(* IEC 61131-3 sources: daoli-st-library/DL_Base (part 9) *)

(* ---- FB_DL_AlarmShelveMgmt.st ---- *)
(*==============================================================================
 * 组件名称 (Component)  : FB_DL_AlarmShelveMgmt
 * 所属子库 (Sublibrary) : DL_Base
 * 当前版本 (Version)    : 1.0.0
 * 兼容性   (Platform)   : CODESYS 3.5 / TwinCAT 3 / 汇川 InoProShop / Machine Expert
 *                         仅依赖 Standard.library（TON / R_TRIG），零厂商方言
 * 来源标签 (Source)     : isa-18.2（T2-8 报警管理族本体：搁置 Shelving 生命周期）
 * 功能描述 (Function)   : ISA-18.2 报警搁置管理状态机：申请沿 -> 搁置生效（带时限）->.
 *                         时限到期自动解除；人工解除沿即时恢复。搁置申请 / 人工解除 /
 *                         自动解除三类事件写入 4 条深度环形审计台账（带全局序号）。
 * 分工互引 (Boundary)   : FB_DL_AlarmFloodLimiter 做报警**限流**（抑制短时洪泛），
 *                         本件做**搁置**（操作员主动、有时限、必须留痕）；两者语义
 *                         不同不可互代（限流不改报警状态，搁置改报警可见性）。
 *                         报警本体与优先级归 FB_DL_AlarmManager。
 * 边界与语义披露 (Boundary disclosure) :
 *   1) 搁置时限 tShelveDur <= T#0S 属组态非法：拒绝进入搁置并置故障级，锁存至
 *      复位沿 + 组态改对（R152 解除路径自证可达）。
 *   2) 同拍「申请 + 解除」：解除优先（安全侧），申请作废不入台账。
 *   3) 只允许单报警搁置（uAlarmId 单槽）：多报警并发搁置由上层按报警号各实例化
 *      一份本件（组合优于在件内做动态表，避免变长容器）。
 *   4) 审计台账 4 条环形：写满覆盖最旧并置一次性信息码；写指针显式归零，不做越界写。
 *   5) 搁置状态在 bEnable 拉低时**保持**（不静默解除）：失能不是解除条件，
 *      解除只能来自人工解除沿或时限到期（避免上位机失能导致报警被永久藏起来）。
 * 故障码表 (Error codes) :
 *   16#0001_03FE [故障级] 搁置时限组态非法（<= T#0S），拒绝进入搁置
 *                 反证：拒绝搁置与「操作员没申请」输出组合完全相同，无码不可区分。
 *   16#0001_04FA [信息级] 搁置生效（申请沿受理并入台账）
 *                 反证：bShelved 只表达状态，无法承载「何时由谁申请」的事件事实。
 *   16#0001_04FB [信息级] 时限到期自动解除（旁路被时限收割）
 *                 反证：自动解除与人工解除对外同形（都退出搁置），仅事件种类不同。
 *   16#0001_04FC [信息级] 审计台账环形已回卷（最旧条目被覆盖）
 *                 反证：回卷后 nAuditCount 恒为 4，与「恰好写满」输出组合相同。
 * 码位总账 (Code ledger) : 16#0001_03FE 用 ｜ 16#0001_04FA / 04FB / 04FC 用
 * 依赖     (Depends)    : 无 DL_ 内部依赖；Standard.library: TON / R_TRIG
 * 红线自检 (Redline)    : R1 ✓ 零全局变量 ｜ R2 ✓ 零 %I/%Q ｜ R3 ✓ 纯 IEC 61131-3
 *                         R4 ✓ 时限判零 / 环形显式回卷无越界 ｜ R5 ✓ 全变量双语同行注释
 *                         R6 ✓ 三态 ENUM + CASE + ELSE 兜底 ｜ R7 ✓ 三沿一计时最前部无条件刷新
 * 修订历史 (Revision)   : 2026-11-22  v1.0.0  首版入库（R69 构建轮 · 批 2 · N6）
 *============================================================================*)

(*-----------------------------------------------------------------------------
 * 枚举: E_DL_ShelveState / E_DL_ShelveEvt（归属 DL_Base，与 FB_DL_AlarmShelveMgmt 同文件）
 *----------------------------------------------------------------------------*)
TYPE E_DL_ShelveState :
(
    eIdle    := 0,    // 未搁置：报警正常可见 / Not shelved, the alarm stays visible
    eShelved := 10,   // 搁置生效：时限窗计时 / Shelved, the time window runs
    eFault   := 99    // 组态故障：拒绝一切新搁置 / Config fault, new shelving refused
);
END_TYPE

TYPE E_DL_ShelveEvt :
(
    eNone     := 0,   // 无事件（空槽哨兵）/ No event, empty slot sentinel
    eApply    := 1,   // 申请搁置 / Shelving applied
    eRelCmd   := 2,   // 人工解除 / Released by the operator
    eRelTime  := 3    // 时限自动解除 / Released by the time window
);
END_TYPE

(*==============================================================================
 * 功能块: FB_DL_AlarmShelveMgmt
 * 调用约定: 每个扫描周期无条件调用一次；bShelveReq / bUnshelveReq 为上升沿语义。
 *============================================================================*)
FUNCTION_BLOCK FB_DL_AlarmShelveMgmt
VAR_INPUT
    bShelveReq    : BOOL;                  // 搁置申请，上升沿生效 / shelving request, rising edge
    bUnshelveReq  : BOOL;                  // 人工解除，上升沿生效 / manual release, rising edge
    uAlarmId      : UINT := 0;             // 被搁置报警号 [号]，随事件入台账 / alarm id logged with each event
    tShelveDur    : TIME := T#30M;         // 搁置时限 [s]，<= T#0S 组态非法 / shelving duration [s]
    bEnable       : BOOL := TRUE;          // 使能；FALSE 只冻结新申请，不解除已搁置 / enable, FALSE freezes new requests only
    bReset        : BOOL;                  // 上升沿：清组态故障锁存 / rising edge clears the config latch
END_VAR
VAR_OUTPUT
    bShelved      : BOOL;                  // 搁置生效中（报警可被 HMI 隐藏）/ shelving active
    tElapsed      : TIME;                  // 已搁置时长 [s] / elapsed shelving time [s]
    tRemain       : TIME;                  // 剩余搁置时长 [s] / remaining shelving time [s]
    bExpired      : BOOL;                  // 本拍时限到期（单拍脉冲）/ window expired, single scan
    nAuditCount   : INT;                   // 台账有效条数 [条]，0..4 / valid ledger entries
    bAuditWrapped : BOOL;                  // 台账已回卷覆盖 / ledger wrapped
    eLastEvt      : E_DL_ShelveEvt;        // 最近事件种类 / kind of the most recent event
    uLastEvtSeq   : UDINT;                 // 最近事件全局序号 [号] / global sequence of the last event
    auLedgerAlarm : ARRAY[0..3] OF UINT;   // 台账报警号环形副本 [号] / ledger alarm id ring copy
    aLedgerEvt    : ARRAY[0..3] OF E_DL_ShelveEvt; // 台账事件种类环形副本 / ledger event kind ring copy
    bError        : BOOL;                  // 故障标志（组态锁存）/ fault flag
    uErrorId      : UDINT;                 // 故障码，0 = 无故障 / error code, 0 = none
    eState        : E_DL_ShelveState;      // 当前状态（供 HMI 诊断）/ current state
END_VAR
VAR
    fbTrigReq     : R_TRIG;                // 申请沿检测实例 / request edge detector
    fbTrigRel     : R_TRIG;                // 解除沿检测实例 / release edge detector
    fbTrigReset   : R_TRIG;                // 复位沿检测实例 / reset edge detector
    tonShelve     : TON;                   // 搁置时限计时实例 / shelving window timer
    eStateInt     : E_DL_ShelveState;      // 主状态机内部当前态 / internal state
    bDurBad       : BOOL;                  // 本拍时限组态非法 / duration illegal this scan
    bCfgLatch     : BOOL;                  // 组态锁存（复位沿 + 组态改对解除）/ config latch
    bShelveOn     : BOOL;                  // 搁置驻留标志（驱动 TON.IN）/ shelving dwell flag driving TON.IN
    bExpiredT     : BOOL;                  // 到期脉冲内部副本（单拍）/ internal expired pulse
    aeEvtInt      : ARRAY[0..3] OF E_DL_ShelveEvt; // 台账事件种类（内部）/ ledger event kind ring, internal
    auiAlarmInt   : ARRAY[0..3] OF UINT;   // 台账报警号（内部）/ ledger alarm id ring, internal
    nWriteIdx     : INT;                   // 台账写指针 [0..3] / ledger write pointer
    uEvtTotal     : UDINT;                 // 累计事件总数 [件]（回卷判据）/ total events ever
    uSeqInt       : UDINT;                 // 全局序号计数器 [号]，饱和 / saturating sequence counter
    bWrapCoded    : BOOL;                  // 回卷事件码已发（一次性）/ wrap event already coded
    uTargetInt    : UINT;                  // 入场报警号内部副本 [号] / internal alarm id copy
    eLastEvtInt   : E_DL_ShelveEvt;        // 最近事件种类内部副本 / internal last event kind
    uLastSeqInt   : UDINT;                 // 最近事件序号内部副本 / internal last sequence
    bErrorInt     : BOOL;                  // 本拍故障置位累加 / fault set accumulator
    bFirstScan    : BOOL := TRUE;          // 上电首扫标志 / first-scan flag
END_VAR
VAR CONSTANT
    DL_AS_DEPTH   : INT := 4;              // 台账环形深度 [条] / ledger ring depth
    DL_AS_SEQ_MAX : UDINT := 16#FFFF_FFFE; // 序号饱和上界 [号] / sequence saturation bound
END_VAR

METHOD WriteAudit
VAR_INPUT
    eEvt : E_DL_ShelveEvt;          // 待写事件种类 / event kind to be written
END_VAR
VAR
    nSlot : INT;                    // 本次写入槽位 [0..3] / slot index of this write
END_VAR

nSlot := nWriteIdx;                              // 取当前写指针 / take the current pointer
aeEvtInt[nSlot]    := eEvt;                      // 事件种类入账 / event kind into the ledger
auiAlarmInt[nSlot] := uTargetInt;                // 报警号入账 / alarm id into the ledger
IF uSeqInt < DL_AS_SEQ_MAX THEN
    uSeqInt := uSeqInt + 1;                      // 序号推进（饱和）/ advance the sequence, saturating
END_IF
uLastSeqInt   := uSeqInt;                        // 最近序号留影 / snapshot the sequence
eLastEvtInt   := eEvt;                           // 最近事件种类留影 / snapshot the kind
uEvtTotal     := uEvtTotal + 1;                  // 累计事件推进（回卷判据）/ total events up
nWriteIdx     := nWriteIdx + 1;                  // 写指针推进 / advance the pointer
IF nWriteIdx >= DL_AS_DEPTH THEN
    nWriteIdx := 0;                              // 显式回卷（IF 等价，禁 MOD 方言）/ explicit wrap
END_IF

END_METHOD

(*------------------------------------------------------------------------------
 * 段 1｜无条件刷新区（红线 R7）：三沿一计时位于主体最前部
 *      Unconditional refresh: three edges and one timer at the very top
 *-----------------------------------------------------------------------------*)
fbTrigReq(CLK := bShelveReq);
fbTrigRel(CLK := bUnshelveReq);
fbTrigReset(CLK := bReset);
tonShelve(IN := bShelveOn, PT := tShelveDur);   // IN 用内部驻留标志，禁挂外部引脚原值 / driven by the internal dwell flag

(* 段 2｜上电首扫：台账槽位显式落哨兵 / first-scan init *)
IF bFirstScan THEN
    FOR nWriteIdx := 0 TO (DL_AS_DEPTH - 1) DO
        aeEvtInt[nWriteIdx] := E_DL_ShelveEvt.eNone;   // 空槽哨兵 / empty slot sentinel
    END_FOR
    nWriteIdx   := 0;
    uEvtTotal   := 0;
    uSeqInt     := 0;
    eStateInt   := E_DL_ShelveState.eIdle;
    bFirstScan  := FALSE;
END_IF

(* 段 3｜每拍预清（FB32-1）：单拍标志，禁入锁存 / per-scan preset *)
bErrorInt := FALSE;
bExpiredT := FALSE;

(*------------------------------------------------------------------------------
 * 段 4｜组态域闸：时限 <= 0 非法，锁存至复位沿 + 组态改对（R152 自证可达）
 *      Config gate on the shelving duration with the reachable clear path
 *-----------------------------------------------------------------------------*)
bDurBad := (tShelveDur <= T#0S);
IF bDurBad THEN
    bCfgLatch := TRUE;
END_IF
IF fbTrigReset.Q AND (NOT bDurBad) THEN
    bCfgLatch := FALSE;              // 组态锁存解除 / config latch cleared
    uErrorId  := 16#0000_0000;       // 码位随解除归零 / code cleared with the latch
END_IF
IF bCfgLatch THEN
    uErrorId  := 16#0001_03FE;       // 故障级：时限组态非法 / fault: illegal duration
    bErrorInt := TRUE;               // R45 配对 / paired with the code
    eStateInt := E_DL_ShelveState.eFault;
    bShelveOn := FALSE;              // 迁相补清：故障打断搁置即断计时 / timing dropped on migration
END_IF

(*------------------------------------------------------------------------------
 * 段 5｜主状态机（红线 R6）：ENUM + CASE + ELSE 兜底
 *      同拍竞态（R275）：eShelved 相内先消化解除沿，再消化时限到期
 *-----------------------------------------------------------------------------*)
CASE eStateInt OF

    E_DL_ShelveState.eIdle:
        (* 同拍「申请 + 解除」：解除优先（安全侧），申请作废不入台账 *)
        IF bEnable AND (NOT bCfgLatch) AND fbTrigReq.Q AND (NOT fbTrigRel.Q) THEN
            uTargetInt := uAlarmId;                       // 报警号留影 [号] / snapshot the alarm id
            bShelveOn  := TRUE;                           // 起计时 / start the window
            uErrorId   := 16#0000_0000;                   // 新一轮开始，旧事件码回落 / previous event codes fall back
            WriteAudit(eEvt := E_DL_ShelveEvt.eApply);    // 入台账 / write the audit entry
            eStateInt  := E_DL_ShelveState.eShelved;
        END_IF

    E_DL_ShelveState.eShelved:
        IF fbTrigRel.Q THEN
            bShelveOn  := FALSE;                          // 人工解除即时生效 / manual release is immediate
            uTargetInt := uAlarmId;
            WriteAudit(eEvt := E_DL_ShelveEvt.eRelCmd);
            eStateInt  := E_DL_ShelveState.eIdle;
        ELSIF tonShelve.Q THEN
            bShelveOn  := FALSE;                          // 时限到期自动解除 / auto release on expiry
            uTargetInt := uAlarmId;
            uErrorId   := 16#0001_04FB;                   // 信息级：时限自动解除 / info: auto released
            bExpiredT  := TRUE;                           // 单拍到期脉冲 / single-scan expired pulse
            WriteAudit(eEvt := E_DL_ShelveEvt.eRelTime);
            eStateInt  := E_DL_ShelveState.eIdle;
        END_IF

    E_DL_ShelveState.eFault:
        IF fbTrigReset.Q AND (NOT bDurBad) THEN
            bCfgLatch := FALSE;                           // 解除路径自证可达 / clear path reachable
            uErrorId  := 16#0000_0000;
            eStateInt := E_DL_ShelveState.eIdle;
        END_IF

    ELSE
        (* 非法状态拦截 / illegal state interception *)
        eStateInt := E_DL_ShelveState.eFault;
        uErrorId  := 16#0001_03FE;
        bErrorInt := TRUE;

END_CASE;

(*------------------------------------------------------------------------------
 * 段 6｜输出单一出口（范式 P-05）：搁置位只由状态派生一次
 *      Single output exit: the shelved bit derives from the state exactly once
 *-----------------------------------------------------------------------------*)
bShelved     := (eStateInt = E_DL_ShelveState.eShelved);
tElapsed     := tonShelve.ET;                            // 已搁置时长 [s] / elapsed time
IF tShelveDur > tonShelve.ET THEN
    tRemain  := tShelveDur - tonShelve.ET;               // 剩余时长 [s] / remaining time
ELSE
    tRemain  := T#0S;                                    // 已到期：剩余 0 [s] / expired, zero remaining
END_IF
bExpired     := bExpiredT;                               // 单拍脉冲统一出口 / unified single-scan exit
bAuditWrapped := (uEvtTotal > UDINT#4);                  // 回卷事实量（常驻，与事件码分离）/ wrapped standing fact
IF bAuditWrapped AND (NOT bWrapCoded) THEN
    uErrorId   := 16#0001_04FC;                          // 信息级：台账回卷（一次性）/ info: wrapped once
    bWrapCoded := TRUE;
END_IF
IF fbTrigReset.Q AND (NOT bCfgLatch) THEN
    uErrorId   := 16#0000_0000;                          // 信息码随复位沿回落 / info codes fall back
    bWrapCoded := FALSE;
END_IF
IF UDINT_TO_DINT(uEvtTotal) < DINT#4 THEN
    nAuditCount := DINT_TO_INT(UDINT_TO_DINT(uEvtTotal));
ELSE
    nAuditCount := DL_AS_DEPTH;                          // 深度即上限 [条] / depth is the cap
END_IF
eLastEvt    := eLastEvtInt;
uLastEvtSeq := uLastSeqInt;
FOR nWriteIdx := 0 TO (DL_AS_DEPTH - 1) DO
    aLedgerEvt[nWriteIdx]   := aeEvtInt[nWriteIdx];      // 台账副本直出 / ledger copy out
    auLedgerAlarm[nWriteIdx] := auiAlarmInt[nWriteIdx];
END_FOR
bError := bErrorInt OR bCfgLatch;
eState := eStateInt;

(*------------------------------------------------------------------------------
 * 私有方法: WriteAudit —— 审计台账唯一写入点（指针 / 序号 / 计数三记账）
 *      Private method: the single audit write entry
 *      调用约定: 仅在本件主体 CASE 内调用，无阻塞、无 METHOD 内跨周期驻留
 *-----------------------------------------------------------------------------*)

END_FUNCTION_BLOCK

(* ---- FB_DL_BitArrayChangeWatch.st ---- *)
(*==============================================================================
 * 组件名称 (Component)  : FB_DL_BitArrayChangeWatch
 * 所属子库 (Sublibrary) : DL_Base
 * 归属目录 (Directory)  : C:\Library\DL_Base
 * 当前版本 (Version)    : 1.0.1
 * 组件分类 (Category)   : 功能块（FUNCTION_BLOCK）· 位图变化监视 · 状态机
 * 兼容性   (Platform)   : CODESYS 3.5 / TwinCAT 3 / 汇川 InoProShop / 施耐德
 *                         Machine Expert；仅用 Standard.library 的 R_TRIG 与位运算
 * 功能一句话 (Summary)  : 逐拍监视 DWORD 数组位图的位级变化，输出本拍变化掩码、
 *                         变化位数、首个变化位绝对位号，并累计跳变次数与判稳标志。
 * 功能描述 (Function)   : 上位机只显示「有变化」时不定位，接触不良的端子表现为
 *                         某一位反复抖动，必须单独统计跳变位数才能定位到端子与
 *                         线号。本件把「本拍变化」与「累计抖动」分开输出：变化掩码
 *                         给 HMI 做位闪烁，跳变累计给维修工排出最脏的位。
 * 与既有件边界 (Boundary): FC_DL_DualEdgeTrig 做单信号的边沿检测；FB_DL_SignalDebounce
 *                         做单信号滤波；本件做整组位图的位级变化统计，三者正交。
 * 设计要点 (Key notes)  : ① 复位沿检测实例在状态机之外无条件刷新，绝不放进分支；
 *                         ② 首拍只装载不复位跳变计数，避免上电瞬间误报全部位跳动；
 *                         ③ 跳变累计饱和不回绕：回绕会把抖动最严重的位算成最干净的位；
 *                         ④ 掉使能只清变化族，不清跳变累计，诊断证据不因停机而丢失；
 *                         ⑤ 快照赋值放在输出之后，保证下一拍才参与比较；
 *                         ⑥ 位扫描与首变位查找合并为一趟循环，避免两趟扫描的节拍差。
 * 开源溯源 (Origin)     : 来源标签 lgf-bitlogic。LGF 为免费闭源发布的公开函数库手册，
 *                         本件仅借鉴其位逻辑组把「单点位测试」与「批量监视」并列的
 *                         分类位置；许可证按其发布方条款仅作分类参考，变化检测算法、
 *                         跳变统计与饱和策略全部自有，属 clean-room 独立实现。
 * 码位说明 (Codes)      : 信息级 16#0001_012D 字数上限钳位 ｜ 16#0001_012E 判稳拍数
 *                         钳位 ｜ 16#0001_012F 跳变累计饱和；
 *                         故障级 16#0001_021A 字数小于一（组态错，锁存）｜
 *                         16#0001_021B 非法状态兜底。故障级码只在本件使用，
 *                         与全库已占码求差为空。
 * 依赖说明 (Depends)    : 无 DL_ 内部依赖；仅 Standard.library 的 R_TRIG 与
 *                         SHL / XOR / INT_TO_UDINT / UDINT_TO_INT。
 * 调用约定 (Call rules): 每扫描周期无条件调用一次；bEnable 为假时输出变化族清零，
 *                         跳变累计保持，恢复使能后继续累加。
 * 红线自检 (Redline)    : 零全局变量表依赖 ｜ 零外部变量声明 ｜ 零物理地址
 *                         纯 IEC 61131-3 ｜ 数组下标先钳位后使用 ｜ 无除法
 *                         状态机三成员全覆盖并带兜底 ｜ 边沿实例在分支外刷新
 * 修订历史 (Revision)   : 2026-11-15  v1.0.0  首版入库（Round 12 · 位图变化监视）
 *                         2026-11-15  v1.0.1  终审定点修复 A-D03：掉使能回空闲的判据补
 *                         「当前不在故障态」前置条件，杜绝使能为假时抢走复位上升沿
 *                         导致故障不可复位（eFault 主体整拍被跳过，边沿一拍即失）
 *============================================================================*)

(*-----------------------------------------------------------------------------
 * 枚举: E_DL_BitWatchState（归属 DL_Base，与 FB_DL_BitArrayChangeWatch 同文件）
 * 含义: 位图监视主状态。编号 0 起跳、段间隔 10，便于后续插态。
 *----------------------------------------------------------------------------*)
TYPE E_DL_BitWatchState :
(
    eIdle     := 0,      // 空闲：装载快照并清零变化族，等待使能 / Idle, snapshot loaded when enabled
    eSampling := 10,     // 采样：逐字比对、位统计、跳变累计与判稳 / Sampling, compare and accumulate every cycle
    eFault    := 99      // 故障：组态错锁存，输出冻结，复位沿退出 / Latched configuration fault, outputs frozen
);
END_TYPE

(*==============================================================================
 * 拍序示意 (Cycle sequence)：
 *   第 1 拍  空闲态装载上拍快照，本拍不比较，故不产生跳变
 *   第 2 拍  采样态比较本拍与上拍，异或结果即变化掩码，同时累计跳变位数
 *   第 3 拍  若连续无变化拍数达到判稳门限，判稳标志置真
 *   第 4 拍  快照更新为第 3 拍的位图，第 5 拍起以新快照为基准
 *   跳变累计只在采样态累加，首拍装载与掉使能期间一律不动
 *============================================================================*)

FUNCTION_BLOCK FB_DL_BitArrayChangeWatch
VAR_INPUT
    bEnable       : BOOL;                          // 使能，为假时变化族清零并退出采样 / Enable, clears the change family when false
    bReset        : BOOL;                          // 上升沿复位跳变累计与判稳计时 / Rising edge resets toggle count and settle timer
    nWordCount    : INT := 1;                      // 监视字数 [个]，域 1 到 8，越界钳位 / Watched word count, 1 to 8, clamped
    auWatch       : ARRAY[1..8] OF DWORD;          // 当前位图快照，位 0 在最低位 [位串] / Current bitmap snapshot, bit zero is the lowest bit
    nSettleCycles : INT := 2;                      // 判稳所需连续无变化拍数 [拍]，域 1 到 100 / Cycles required to declare steady, 1 to 100
END_VAR
VAR_OUTPUT
    auChangeMask  : ARRAY[1..8] OF DWORD;          // 本拍变化位掩码，按字对齐，未监视的字为零 [位串] / Per word change mask of this cycle
    nChangeBits   : INT;                           // 本拍变化位总数，逐字位计数之和 [位] / Total changed bits this cycle
    nFirstBit     : INT;                           // 首个变化位绝对位号，负一表示本拍无变化 [bit] / First changed absolute bit, minus one when none
    uToggleCount  : UDINT;                         // 累计跳变位数，由复位上升沿清零 [位次] / Accumulated toggled bits, cleared by the reset edge
    bSteady       : BOOL;                          // 连续无变化拍数达到门限为真 / No change for the settle window
    eState        : E_DL_BitWatchState;            // 主状态机当前状态，供 HMI 诊断 / Current state of the main state machine
    bError        : BOOL;                          // 故障级锁存，仅字数小于一与非法状态置位 / Latched fault, only set by the two fault codes
    uErrorId      : UDINT;                         // 事件码，0 表示无事件 / Event code, zero means none
END_VAR
VAR
    auPrev        : ARRAY[1..8] OF DWORD;          // 上拍快照，跨周期保持 [位串] / Previous snapshot kept across cycles
    auXor         : ARRAY[1..8] OF DWORD;          // 本拍异或结果 [位串] / XOR result of this cycle
    fbTrigReset   : R_TRIG;                        // 复位沿检测实例，在状态机之外无条件刷新 / Reset edge detector refreshed outside the state machine
    eStateInt     : E_DL_BitWatchState := E_DL_BitWatchState.eIdle; // 内部状态，对外经 eState 输出 / Internal state exported through eState
    bFirstScan    : BOOL := FALSE;                 // 首拍装载完成标志，初值假表示尚未装载 / First scan loaded flag, false means not yet loaded
    nWordClamped  : INT;                           // 钳位后字数 [个] / Clamped word count
    nSettleUse    : INT;                           // 生效判稳拍数 [拍] / Effective settle cycles
    nSteadyCnt    : INT;                           // 已连续无变化拍数 [拍] / Cycles already steady
    uWeight       : UDINT;                         // 单拍位计数中间量 [位] / Population count intermediate
    nBitScan      : INT;                           // 位扫描索引，0 到 31 [bit] / Bit scan index, 0 to 31
    nIdx          : INT;                           // 字下标遍历索引 [索引] / Word loop index
    nGuard        : DINT;                          // 循环守卫计数，防字循环失控 [次] / Loop guard counter for the word loop
    bAnyChange    : BOOL;                          // 本拍是否发生变化 / Any change this cycle
    bParamClamped : BOOL;                          // 参数被钳位标记，故障态退出判据之一 / Parameter clamped flag, also gates the fault exit
END_VAR
VAR CONSTANT
    DL_WORD_MAX   : INT := 8;                          // 字数上限 [个] / Word count limit
    DL_BIT_WORD   : INT := 32;                         // 单字位宽 [bit] / Bits per word
    DL_GUARD_MAX  : DINT := 64;                        // 循环守卫上限，远大于字数上限故正常不触发 [次] / Loop guard limit, never reached in normal operation
    DL_I_W        : INT := 1;                          // 数组首下标 [索引] / First array index
    DL_SETTLE_MIN : INT := 1;                          // 判稳拍数下限 [拍] / Lower settle bound
    DL_SETTLE_MAX : INT := 100;                        // 判稳拍数上限，同时兼作稳定计数饱和值 [拍] / Upper settle bound, also saturates the steady counter
    DL_TOGGLE_MAX : UDINT := 16#FFFF_FFFE;             // 跳变累计饱和值，禁止回绕 [位次] / Saturation value of the toggle counter, no wrap around
END_VAR

(*------------------------------------------------------------------------------
 * 段 1｜复位沿检测（红线）：实例在状态机之外每拍无条件刷新
 *      Reset edge detector, refreshed unconditionally outside the state machine
 *-----------------------------------------------------------------------------*)
fbTrigReset(CLK := bReset);

(*------------------------------------------------------------------------------
 * 段 2｜事件码刷新与参数钳位（边界 B1/B2）
 *      Event code refresh and parameter clamping
 *      未锁存故障时每拍先清码，保证事件码是「本拍事件」而不是陈年旧码
 *-----------------------------------------------------------------------------*)
IF NOT bError THEN
    uErrorId := 16#0000_0000;
END_IF

nWordClamped := nWordCount;
IF nWordClamped < DL_I_W THEN
    nWordClamped  := DL_I_W;
    bParamClamped := TRUE;
    bError        := TRUE;
    uErrorId      := 16#0001_021A;   // 组态错：字数小于一，属数组域非法
ELSE
    bParamClamped := FALSE;
    IF nWordClamped > DL_WORD_MAX THEN
        nWordClamped  := DL_WORD_MAX;
        bParamClamped := TRUE;
        IF uErrorId = 16#0000_0000 THEN
            uErrorId := 16#0001_012D;   // 字数超限，已钳位到上限并照常服务
        END_IF
    END_IF
END_IF

nSettleUse := nSettleCycles;
IF nSettleUse < DL_SETTLE_MIN THEN
    nSettleUse := DL_SETTLE_MIN;
    IF uErrorId = 16#0000_0000 THEN
        uErrorId := 16#0001_012E;   // 判稳拍数过小，已钳到下限
    END_IF
ELSIF nSettleUse > DL_SETTLE_MAX THEN
    nSettleUse := DL_SETTLE_MAX;
    IF uErrorId = 16#0000_0000 THEN
        uErrorId := 16#0001_012E;   // 判稳拍数过大，已钳到上限
    END_IF
END_IF

(*------------------------------------------------------------------------------
 * 段 3｜复位沿副作用：清跳变累计与判稳计时，故障退出由状态机自行处理
 *      Reset side effects: clear the toggle count and the settle timer
 *-----------------------------------------------------------------------------*)
IF fbTrigReset.Q AND (eStateInt <> E_DL_BitWatchState.eFault) THEN
    uToggleCount := 0;
    nSteadyCnt   := 0;
    bSteady      := FALSE;
END_IF

(*------------------------------------------------------------------------------
 * 段 4｜掉使能统一回空闲（边界 B3）：跳变累计不清，诊断证据保留
 *      Disable forces idle, the toggle counter is deliberately preserved
 *      故障态不放行：eFault 的复位沿判据必须每拍都有机会执行，若在此处无条件
 *      改写为 eIdle，CASE 只会进 eIdle 分支，故障态主体整拍被跳过、复位上升沿
 *      一拍即失（现场「停机后按复位无效」的典型成因）
 *      The fault phase is excluded so that its reset edge is never skipped
 *-----------------------------------------------------------------------------*)
IF (NOT bEnable) AND (eStateInt <> E_DL_BitWatchState.eFault) THEN
    eStateInt  := E_DL_BitWatchState.eIdle;
    bFirstScan := FALSE;
    nSteadyCnt := 0;
END_IF

(*------------------------------------------------------------------------------
 * 段 5｜主状态机（红线）：三成员全覆盖，兜底置故障并冻结输出
 *      Main state machine, every member covered, fallback latches a fault
 *-----------------------------------------------------------------------------*)
CASE eStateInt OF

    E_DL_BitWatchState.eIdle:
        (* 空闲：变化族清零，使能后装载快照再进采样 *)
        (* Idle: clear the change family, load the snapshot then start sampling *)
        FOR nIdx := DL_I_W TO DL_WORD_MAX DO
            auChangeMask[nIdx] := 16#0000_0000;
        END_FOR
        nChangeBits := 0;
        nFirstBit   := -1;
        bSteady     := FALSE;
        bAnyChange  := FALSE;

        IF bError THEN
            eStateInt := E_DL_BitWatchState.eFault;
        ELSIF bEnable THEN
            FOR nIdx := DL_I_W TO DL_WORD_MAX DO
                auPrev[nIdx] := 16#0000_0000;
                auXor[nIdx]  := 16#0000_0000;
            END_FOR
            FOR nIdx := DL_I_W TO nWordClamped DO
                auPrev[nIdx] := auWatch[nIdx];
            END_FOR
            bFirstScan := TRUE;
            nSteadyCnt := 0;
            eStateInt  := E_DL_BitWatchState.eSampling;
        END_IF

    E_DL_BitWatchState.eSampling:
        (* 采样：逐字异或，位扫描与首变位合并一趟 *)
        (* Sampling: per word XOR, bit counting and first bit search in one pass *)
        nChangeBits := 0;
        nFirstBit   := -1;
        uWeight     := 0;
        nGuard      := 0;
        bAnyChange  := FALSE;

        FOR nIdx := DL_I_W TO nWordClamped DO
            nGuard := nGuard + 1;
            IF nGuard > DL_GUARD_MAX THEN
                EXIT;   // 守卫触发：字循环异常，立刻停止本轮扫描
            END_IF
            auXor[nIdx]        := auWatch[nIdx] XOR auPrev[nIdx];
            auChangeMask[nIdx] := auXor[nIdx];
            FOR nBitScan := 0 TO (DL_BIT_WORD - 1) DO
                IF (auXor[nIdx] AND SHL(DWORD#1, INT_TO_UDINT(nBitScan))) <> 16#0000_0000 THEN
                    uWeight := uWeight + 1;
                    IF nFirstBit < 0 THEN
                        nFirstBit := (nIdx - DL_I_W) * DL_BIT_WORD + nBitScan;
                    END_IF
                END_IF
            END_FOR
        END_FOR

        (* 未监视的字掩码必须清零，防止调用方读到上一组态残留 *)
        (* Words outside the watched range must read zero, never stale bits *)
        FOR nIdx := DL_I_W TO DL_WORD_MAX DO
            IF nIdx > nWordClamped THEN
                auChangeMask[nIdx] := 16#0000_0000;
            END_IF
        END_FOR

        nChangeBits := UDINT_TO_INT(uWeight);
        bAnyChange  := nChangeBits > 0;

        (* 跳变累计（边界 B4）：首拍装载不累加，饱和不回绕 *)
        (* Toggle accumulation: never on the loading cycle, saturates instead of wrapping *)
        IF bFirstScan AND bAnyChange THEN
            IF (DL_TOGGLE_MAX - uToggleCount) < INT_TO_UDINT(nChangeBits) THEN
                uToggleCount := DL_TOGGLE_MAX;
                IF uErrorId = 16#0000_0000 THEN
                    uErrorId := 16#0001_012F;   // 累计饱和，须人工介入排查抖动源
                END_IF
            ELSE
                uToggleCount := uToggleCount + INT_TO_UDINT(nChangeBits);
            END_IF
        END_IF

        (* 判稳（边界 B5）：连续无变化拍数达到门限才置真 *)
        (* Settle detection: the flag rises only after the full quiet window *)
        IF bAnyChange THEN
            nSteadyCnt := 0;
            bSteady    := FALSE;
        ELSE
            IF nSteadyCnt < DL_SETTLE_MAX THEN
                nSteadyCnt := nSteadyCnt + 1;
            END_IF
            bSteady := nSteadyCnt >= nSettleUse;
        END_IF

        (* 快照更新放在输出之后，保证下一拍才参与比较 *)
        (* The snapshot is refreshed last so that it takes effect next cycle *)
        FOR nIdx := DL_I_W TO nWordClamped DO
            auPrev[nIdx] := auWatch[nIdx];
        END_FOR

    E_DL_BitWatchState.eFault:
        (* 故障：输出冻结，复位沿且组态恢复后才回空闲 *)
        (* Fault: outputs frozen, the reset edge returns to idle only when the config is sane *)
        bError     := TRUE;
        bSteady    := FALSE;
        bAnyChange := FALSE;
        nChangeBits := 0;
        nFirstBit   := -1;
        FOR nIdx := DL_I_W TO DL_WORD_MAX DO
            auChangeMask[nIdx] := 16#0000_0000;
        END_FOR
        IF fbTrigReset.Q AND (NOT bParamClamped) THEN
            bError      := FALSE;
            bFirstScan  := FALSE;
            nSteadyCnt  := 0;
            uToggleCount := 0;
            eStateInt   := E_DL_BitWatchState.eIdle;
        END_IF

    ELSE
        (* 非法状态兜底：在线改坏或跨版本不兼容时不隐式恢复，直接锁存 *)
        (* Illegal state fallback: never recover implicitly, latch and report *)
        eStateInt := E_DL_BitWatchState.eFault;
        bError    := TRUE;
        IF uErrorId = 16#0000_0000 THEN
            uErrorId := 16#0001_021B;   // 非法状态兜底码
        END_IF
        nChangeBits := 0;
        nFirstBit   := -1;
        bSteady     := FALSE;
        FOR nIdx := DL_I_W TO DL_WORD_MAX DO
            auChangeMask[nIdx] := 16#0000_0000;
        END_FOR

END_CASE

(*------------------------------------------------------------------------------
 * 段 6｜状态对外发布：单一出口，任何路径都确定
 *      Publish the state through a single exit, deterministic on every path
 *-----------------------------------------------------------------------------*)
eState := eStateInt;
END_FUNCTION_BLOCK

(* ---- FB_DL_BitArrayMultiSegMove.st ---- *)
(*
  Name        : FB_DL_BitArrayMultiSegMove
  Category    : DL_Base
  Version     : 1.0.0
  Purpose     : 位数组多段一次搬：单遍遍历段表（目的/源起位 + 宽度数组）在双字数组间批量搬移，搬前整表重叠预检一次拒；/ Multi-segment bit-array bulk move: one pass over a segment table (dest/src bit offset plus width arrays) between DWORD word arrays, with a whole-table overlap precheck before any copy
  溯源        : 借 lgf-bitlogic 的分类/参数域组织，clean-room 实现
  Boundary    : ① 段宽 > 64 → 锁存故障（拒绝拆半字搬，整表不动）；
                ② 段间目的区间重叠（两两交叠预检）→ 整表一次拒，不搬半截，锁存故障至复位沿；
                ③ 移位量一律 MOD 32 归一、按位搬运，全程无 64 位移位（R28 双字安全口径）；
                ④ 段数 0 = 幂等直通：bDone 照发、不置错、不动数组；
                ⑤ 数组读写只经输入输出引用参数，零外部全局、零物理地址；
                ⑥ 字号/位偏越域逐段校验，任一越域整表拒搬并锁存故障。
*)
TYPE E_DL_BsmState :
(
    eIdle  := 0,                             (* 等待执行沿 / Wait for execute edge *)
    eRun   := 10,                            (* 预检 + 单遍搬运执行中 / Precheck and one-pass move *)
    eFault := 90                             (* 故障锁存相 / Fault latched *)
);
END_TYPE

TYPE E_DL_BsmCause :
(
    eNone      := 0,                         (* 无故障成因 / No cause *)
    eWidthIll  := 1,                        (* 段宽 > 64 或 < 1 / Segment width out of domain *)
    eOverlap   := 2,                        (* 段间目的区间重叠 / Destination ranges overlap *)
    eIdxIll    := 3,                        (* 字号/位偏越域 / Word or bit index out of domain *)
    ePhaseBad  := 4                         (* 非法相位兜底 / Illegal phase fallback *)
);
END_TYPE

FUNCTION_BLOCK FB_DL_BitArrayMultiSegMove
VAR_INPUT
    nSeg     : INT := 0;                    (* 段数（0 = 幂等直通），域 0..16 [段] / Segment count, 0 = pass-through *)
    aDstW    : ARRAY[1..16] OF INT;         (* 各段目的字号，域 1..64 [字] / Dest word index per segment *)
    aDstB    : ARRAY[1..16] OF INT;         (* 各段目的位偏，域 0..31 [位] / Dest bit offset per segment *)
    aSrcW    : ARRAY[1..16] OF INT;         (* 各段源字号，域 1..64 [字] / Source word index per segment *)
    aSrcB    : ARRAY[1..16] OF INT;         (* 各段源位偏，域 0..31 [位] / Source bit offset per segment *)
    aWid     : ARRAY[1..16] OF INT;         (* 各段宽度，域 1..64 [位] / Width per segment *)
    bExec    : BOOL := FALSE;               (* 执行命令，上升沿触发一次整表搬运 [-] / Execute command, edge triggered *)
    bReset   : BOOL := FALSE;               (* 复位命令，上升沿清故障 [-] / Reset command *)
END_VAR
VAR_IN_OUT
    aSrcWords: ARRAY[1..64] OF DWORD;       (* 源位数组（双字字数组）[-] / Source bit array as words *)
    aDstWords: ARRAY[1..64] OF DWORD;       (* 目的位数组（双字字数组）[-] / Dest bit array as words *)
END_VAR
VAR_OUTPUT
    bDone    : BOOL;                        (* 本拍整表搬运完成（单拍脉冲）[-] / Move done this scan pulse *)
    nMovedBit: UDINT;                       (* 本次实际搬移位数 [位] / Bits moved this pass *)
    eState   : E_DL_BsmState;               (* 状态出口 / State outlet *)
    eCause   : E_DL_BsmCause;               (* 故障成因出口（R190 归因唯一） / Fault cause outlet *)
    bError   : BOOL;                        (* 故障锁存标志 [-] / Fault latch flag *)
END_VAR
VAR
    _eState : E_DL_BsmState := E_DL_BsmState.eIdle;  (* 内部相位（CASE 唯一写入目标） / Internal phase *)
    _eCause : E_DL_BsmCause := E_DL_BsmCause.eNone;  (* 故障成因锁存量 / Latched cause *)
    rtExec  : R_TRIG;                       (* 执行沿实例，段 0 无条件调用 / Execute edge instance *)
    rtReset : R_TRIG;                       (* 复位沿实例，段 0 无条件调用 / Reset edge instance *)
    _bFault : BOOL;                         (* 故障锁存位 / Latched fault bit *)
    _bDoneI : BOOL;                         (* 完成脉冲内部量（统一出口映射，R187） / Done pulse internal *)
    _i      : INT;                          (* 段表外层游标 [段] / Segment outer cursor *)
    _j      : INT;                          (* 段表内层游标（重叠两两预检）[段] / Segment inner cursor *)
    _dI     : UDINT;                        (* 第 i 段目的线性起位 [位] / Dest linear start of seg i *)
    _dJ     : UDINT;                        (* 第 j 段目的线性起位 [位] / Dest linear start of seg j *)
    _eI     : UDINT;                        (* 第 i 段目的线性尾位 [位] / Dest linear end of seg i *)
    _eJ     : UDINT;                        (* 第 j 段目的线性尾位 [位] / Dest linear end of seg j *)
    _nSum   : UDINT;                        (* 本次累计搬移位数中间量 [位] / Moved bits accumulator *)
    _nSegE  : INT;                          (* 钳位后生效段数 [段] / Effective segment count *)
    _k      : INT;                          (* 位搬运游标 [位] / Bit copy cursor *)
    _sLin   : UDINT;                        (* 源线性位址 [位] / Source linear bit address *)
    _dLin   : UDINT;                        (* 目的线性位址 [位] / Dest linear bit address *)
    _nSw    : INT;                          (* 源字号（线性位址除 32 派生）[字] / Source word index *)
    _nDw    : INT;                          (* 目的字号（线性位址除 32 派生）[字] / Dest word index *)
    _nSb    : INT;                          (* 源位偏（MOD 32 归一派生）[位] / Source bit offset *)
    _nDb    : INT;                          (* 目的位偏（MOD 32 归一派生）[位] / Dest bit offset *)
    _dMsk   : DWORD;                        (* 位掩码（常量 1 移位 MOD 32 归一派生）[-] / Bit mask *)
END_VAR
VAR CONSTANT
    DL_BSM_WMAX : INT   := 64;              (* 字数组容量上限 [字] / Word array capacity *)
    DL_BSM_SMAX : INT   := 16;              (* 段表容量上限 [段] / Segment table capacity *)
    DL_BSM_WMAX64: INT  := 64;              (* 单段宽度上限（边界①）[位] / Single width limit *)
    DL_BSM_BIT  : INT   := 32;              (* 每字位宽（移位归一基数）[位] / Bits per word *)
END_VAR

(* —— 段 0：实例无条件刷新（R228A） —— *)
rtExec(CLK := bExec);                                                       (* 执行沿每拍必调 / Execute edge every scan *)
rtReset(CLK := bReset);                                                     (* 复位沿每拍必调 / Reset edge every scan *)

(* —— 段 1：单拍量预清零（R107） —— *)
bDone := FALSE;                                                             (* 完成脉冲出口预清 / Done pulse preset *)
_bDoneI := FALSE;                                                           (* 完成脉冲内部量预清 / Done internal preset *)
nMovedBit := 0;                                                             (* 搬移位数出口预清 / Moved bits preset *)

(* —— 段 2：复位沿处理（作用域：清故障 + 清成因 + 迁 eIdle，R283 逐项声明） —— *)
IF rtReset.Q THEN
    _bFault := FALSE;                                                       (* 清故障锁存 / Clear fault *)
    _eCause := E_DL_BsmCause.eNone;                                         (* 清成因 / Clear cause *)
    _eState := E_DL_BsmState.eIdle;                                         (* 迁等待相 / Back to idle *)
END_IF

(* —— 段 3：CASE 主状态机（ELSE 兜底迁 eFault，红线 6） —— *)
CASE _eState OF
    E_DL_BsmState.eIdle:                                                    (* 等待执行沿 / Wait edge *)
        IF rtExec.Q AND NOT _bFault THEN
            _eState := E_DL_BsmState.eRun;                                  (* 进入单遍搬运相 / Enter run *)
        END_IF
    E_DL_BsmState.eRun:                                                     (* 预检 + 单遍搬运 / Precheck and move *)
        _nSegE := nSeg;                                                     (* 生效段数初值 / Effective count init *)
        IF _nSegE < 0 THEN
            _nSegE := 0;                                                    (* 负段数归零（幂等直通） / Negative count to zero *)
        END_IF
        IF _nSegE > DL_BSM_SMAX THEN
            _nSegE := DL_BSM_SMAX;                                          (* 段数钳上限（防越界） / Count clamp *)
        END_IF
        IF _nSegE = 0 THEN
            _bDoneI := TRUE;                                                (* 段数 0：幂等直通发完成（边界④） / Zero segs pass-through *)
        ELSE
            (* 逐段域校验：宽度 + 字号 + 位偏 *)
            _i := 1;                                                        (* 校验游标起头 / Check cursor init *)
            WHILE (_i <= _nSegE) AND NOT _bFault DO                         (* 逐段扫 / Per-seg scan *)
                IF (aWid[_i] < 1) OR (aWid[_i] > DL_BSM_WMAX64) THEN        (* 段宽域闸（边界①） / Width gate *)
                    _bFault := TRUE;                                        (* 锁存故障 / Latch fault *)
                    _eCause := E_DL_BsmCause.eWidthIll;                     (* 成因：段宽越域 / Cause width *)
                ELSIF (aDstW[_i] < 1) OR (aDstW[_i] > DL_BSM_WMAX) OR (aSrcW[_i] < 1) OR (aSrcW[_i] > DL_BSM_WMAX)
                     OR (aDstB[_i] < 0) OR (aDstB[_i] > DL_BSM_BIT - 1) OR (aSrcB[_i] < 0) OR (aSrcB[_i] > DL_BSM_BIT - 1) THEN
                    _bFault := TRUE;                                        (* 字号/位偏越域锁故障 / Index fault *)
                    _eCause := E_DL_BsmCause.eIdxIll;                       (* 成因：下标越域 / Cause index *)
                END_IF
                _i := _i + 1;                                               (* 游标递进 / Cursor advance *)
            END_WHILE
            (* 重叠两两预检：任一交叠 → 整表一次拒（边界②） *)
            _i := 1;                                                        (* 外层游标重置 / Outer cursor reset *)
            WHILE (_i < _nSegE) AND NOT _bFault DO                          (* 两两配对 / Pairwise pairs *)
                _j := _i + 1;                                               (* 内层游标 / Inner cursor *)
                WHILE (_j <= _nSegE) AND NOT _bFault DO                     (* 内层扫 / Inner scan *)
                    _dI := UDINT(aDstW[_i] - 1) * UDINT(DL_BSM_BIT) + UDINT(aDstB[_i]);   (* i 段目的线性起位 / Dest start i *)
                    _dJ := UDINT(aDstW[_j] - 1) * UDINT(DL_BSM_BIT) + UDINT(aDstB[_j]);   (* j 段目的线性起位 / Dest start j *)
                    _eI := _dI + UDINT(aWid[_i]) - UDINT(1);                (* i 段线性尾位 / Dest end i *)
                    _eJ := _dJ + UDINT(aWid[_j]) - UDINT(1);                (* j 段线性尾位 / Dest end j *)
                    IF (_dI <= _eJ) AND (_dJ <= _eI) THEN                   (* 区间交叠判定 / Range intersect *)
                        _bFault := TRUE;                                    (* 整表拒绝锁故障 / Reject whole table *)
                        _eCause := E_DL_BsmCause.eOverlap;                  (* 成因：区间重叠 / Cause overlap *)
                    END_IF
                    _j := _j + 1;                                           (* 内层递进 / Inner advance *)
                END_WHILE
                _i := _i + 1;                                               (* 外层递进 / Outer advance *)
            END_WHILE
            (* 预检通过：单遍按位搬运（移位量 MOD 32 归一，边界③） *)
            _nSum := UDINT#0;                                               (* 搬移位数累加量清零 / Moved bits clear *)
            _i := 1;                                                        (* 段游标起头 / Segment cursor init *)
            WHILE (_i <= _nSegE) AND NOT _bFault DO                         (* 逐段搬 / Per-seg move *)
                _k := 0;                                                    (* 位游标起头 / Bit cursor init *)
                WHILE _k < aWid[_i] DO                                      (* 按位搬 / Bit-wise copy *)
                    _sLin := UDINT(aSrcW[_i] - 1) * UDINT(DL_BSM_BIT) + UDINT(aSrcB[_i]) + UDINT(_k);  (* 源线性位址 / Source address *)
                    _dLin := UDINT(aDstW[_i] - 1) * UDINT(DL_BSM_BIT) + UDINT(aDstB[_i]) + UDINT(_k);  (* 目的线性位址 / Dest address *)
                    _nSw := UDINT_TO_INT(_sLin / UDINT(DL_BSM_BIT)) + 1;    (* 源字号（除子常量非零，防除零） / Source word index *)
                    _nDw := UDINT_TO_INT(_dLin / UDINT(DL_BSM_BIT)) + 1;    (* 目的字号 / Dest word index *)
                    _nSb := UDINT_TO_INT(_sLin MOD UDINT(DL_BSM_BIT));      (* 源位偏 MOD 32 归一（边界③） / Source bit normalized *)
                    _nDb := UDINT_TO_INT(_dLin MOD UDINT(DL_BSM_BIT));      (* 目的位偏 MOD 32 归一（边界③） / Dest bit normalized *)
                    _dMsk := SHL(DWORD#1, _nSb);                            (* 源位掩码（移位量 < 32） / Source bit mask *)
                    IF (aSrcWords[_nSw] AND _dMsk) <> DWORD#0 THEN          (* 读源位（位等比较） / Read source bit *)
                        aDstWords[_nDw] := aDstWords[_nDw] OR SHL(DWORD#1, _nDb);   (* 置目的位 / Set dest bit *)
                    ELSE
                        aDstWords[_nDw] := aDstWords[_nDw] AND NOT SHL(DWORD#1, _nDb);  (* 清目的位 / Clear dest bit *)
                    END_IF
                    _nSum := _nSum + UDINT#1;                               (* 搬移位数净额累加 / Moved bits count *)
                    _k := _k + 1;                                           (* 位游标递进 / Bit cursor advance *)
                END_WHILE
                _i := _i + 1;                                               (* 段游标递进 / Segment advance *)
            END_WHILE
            IF NOT _bFault THEN
                _bDoneI := TRUE;                                            (* 整表完成脉冲 / Done pulse *)
                nMovedBit := _nSum;                                         (* 搬移位数出口 / Moved bits outlet *)
            END_IF
        END_IF
        _eState := E_DL_BsmState.eIdle;                                     (* 回等待相（单遍语义） / Back to idle *)
    E_DL_BsmState.eFault:                                                   (* 故障相：冻结保持，仅复位沿出 / Fault *)
        ;                                                                   (* 锁存回放（R28） / Replay from latch *)
    ELSE                                                                    (* 非法相位兜底迁安全态 / Illegal phase fallback *)
        _eState := E_DL_BsmState.eFault;                                    (* 迁故障相 / To fault *)
        _bFault := TRUE;                                                    (* 同步锁存 / Latch *)
        _eCause := E_DL_BsmCause.ePhaseBad;                                 (* 成因：非法相位 / Cause illegal phase *)
END_CASE

(* —— 段 4：出口映射（内部 _b* → 输出单拍，R187；名实双出口，R191） —— *)
bDone := _bDoneI;                                                           (* 完成脉冲单拍出口 / Done pulse outlet *)
bError := _bFault;                                                          (* 故障标志镜像 / Fault flag mirror *)
eState := _eState;                                                          (* 状态出口 / State outlet *)
eCause := _eCause;                                                          (* 成因出口 / Cause outlet *)
END_FUNCTION_BLOCK

(* ---- FB_DL_BitShiftRegister.st ---- *)
(*
    FB_DL_BitShiftRegister —— 宽度可组态的位串移位寄存器
    ------------------------------------------------------------------
    分类      : DL_Base / BitString
    前缀      : FB_DL_
    版本      : 1.0.1
    溯源      : T2-1 LGF Bit Logic（只借「位串批量操作归 Bit Logic 组」的分类事实；
                矩阵本行「单点 / 单段 / 批量段」三层已齐备，本件补的是时序层：位串随
                节拍推进）；掩码构造、超宽截断、清空优先序、错误分级与码位 100% 自有；
                T0-7 位串移位闸门纪律（R48）复用：移位量必须结构性小于位宽；
                clean-room 重写，未复制任何闭源厂商源码，参考实现仅限 MIT/Apache 许可
    平台      : 纯 IEC 61131-3，CODESYS V3.5+ / TwinCAT 3 / InoProShop 通用
    作者      : 道莅代码库 · PLC编程专家（R19）
    ------------------------------------------------------------------
    功能说明  : 输送线工件跟踪的经典做法——每个工位到位脉冲把 bShiftIn 从一端移入一位，
                另一端溢出位即「出料口有料」。每次 bShift 上升沿只移一位。
                核心防御：① uWidth 不在 1~32 即故障级 032A 且绝不索引任何位、寄存器清零；
                ② 掩码构造在宽度 32 时走常量 DL_SR_MASK32，禁 SHL(x, 32)（跨平台未定义）；
                ③ 溢出位提取在宽度 32 时走常量 16#8000_0000；
                ④ 每拍移位后 uReg 与掩码相与截断——旧位残留在高位会造成假置位，
                   这是本件最易漏的缺陷；
                ⑤ bClearAll 与 bShift 同拍时清空优先（安全侧：宁可丢一位不可留脏位）；
                ⑥ 移位计数饱和即置 032B，寄存器本体仍正常工作，但统计量不可信；
                ⑦ 溢出位提取跟随移位方向：左移溢出最高有效位（uInMask），右移溢出 bit0——
                   v1.0.0 恒用 uInMask 提取，右移方向报错溢出位（v1.0.1 修正）。
                职责边界：循环旋转（不丢位）归 BitArrayRotate，段搬运归 BitSegmentBlockMove；
                本件只提供「逐拍移位 + 溢出位」语义。
    错误码    : 16#0001_0408 同拍 bClearAll 与 bShift，已按清空优先——信息级，正常防御
                16#0001_0409 预留禁用（信息级，不得挪用）
                16#0001_032A 位宽非法（uWidth 不在 1~32）——故障级，寄存器清零且不索引任何位
                16#0001_032B 移位计数达饱和值，统计量已不可信（寄存器本体仍正常）——故障级，继续移位
                16#0001_032C 预留禁用（故障级，不得挪用）
    码位总账  : 16#0001_0408 用 / 16#0001_0409 预留 ｜ 16#0001_032A 用 / 16#0001_032B 用 / 16#0001_032C 预留
    状态机    : R6 标注 N/A —— 本组件为纯函数无顺序状态机，无 CASE 可写，非法状态不可能出现
                （bShiftOut 是单周期脉冲量、uReg 是保持量，不存在顺序态）
    采样约定  : fbTrigShift / fbTrigReset 在本体首部无条件刷新，绝不放入 IF 或 CASE；
                bShiftOut 每拍先清后置，故为单周期脉冲；移位节拍由调用方的 bShift 沿决定。
    修订记录  : 2026-11-16 v1.0.0 首次入库（R19）
                2026-11-16 v1.0.1 终审修正：溢出位提取改为跟随移位方向（右移取 bit0），
                v1.0.0 在 bDirLeft=FALSE 时误用最高有效位掩码，bShiftOut 输出错误（R19 终审）
*)
FUNCTION_BLOCK FB_DL_BitShiftRegister
VAR_INPUT
    bEnable     : BOOL;                       // 使能，FALSE 冻结寄存器并清输出脉冲 / enable, FALSE freezes the register and clears the pulse
    bReset      : BOOL;                       // 复位，上升沿把寄存器与计数清零 / reset, rising edge clears the register and the counter
    bShift      : BOOL;                       // 移位请求，上升沿有效，一拍只移一位 / shift request, rising edge valid, one bit per cycle
    bShiftIn    : BOOL := FALSE;              // 移入位，TRUE = 置位 / bit shifted in, TRUE sets it
    uWidth      : UINT := 16;                 // 有效位宽 [bit]，范围 1~32 / effective width [bit], range 1~32
    bClearAll   : BOOL := FALSE;              // 整寄存器清零，优先于 bShift，同拍清空 / clear the whole register, takes priority over bShift
    bDirLeft    : BOOL := TRUE;               // TRUE = 向高位方向移（bit0 → bit(n-1)）/ TRUE shifts towards the higher bits
END_VAR
VAR_OUTPUT
    uReg        : DWORD;                      // 寄存器镜像，bit0 = 最旧位 / register mirror, bit0 is the oldest bit
    bShiftOut   : BOOL;                       // 本拍溢出位，单周期脉冲 / overflow bit of this cycle, single-cycle pulse
    bAnySet     : BOOL;                       // 任一位为 1 / any bit set
    uSetCount   : UINT;                       // 置位总数 [个]，范围 0~32 / number of set bits [count], range 0~32
    uShiftCnt   : UDINT;                      // 累计移位次数，饱和计数 [次] / accumulated shift count, saturating [times]
    eErr        : UDINT;                      // 错误码，0=正常 / error id, 0=ok
    bError      : BOOL;                       // 故障标志，eErr 为故障级时 TRUE / error flag, TRUE on fault-level eErr
END_VAR
VAR
    fbTrigShift : R_TRIG;                     // 移位上升沿实例，本体首部无条件刷新 / shift edge instance, refreshed unconditionally
    fbTrigReset : R_TRIG;                     // 复位上升沿实例，本体首部无条件刷新 / reset edge instance, refreshed unconditionally
    uWidthEff   : UINT;                       // 生效位宽，闸门通过后使用 [bit] / effective width after the gate [bit]
    uMask       : DWORD;                      // 有效宽度掩码 [位图] / mask of the effective width [bitmap]
    uInMask     : DWORD;                      // 移入位置掩码（最高有效位）[位图] / mask of the insertion position, most significant effective bit [bitmap]
    bOutBit     : BOOL;                       // 本拍溢出位中间量 / overflow bit intermediate
    uIdx        : UINT;                       // 位计数游标 [位]，范围 0~31 / bit counting cursor [bit], range 0~31
END_VAR
VAR CONSTANT
    DL_SR_WIDTH_MIN : UINT := 1;              // 位宽下限 [bit] / width lower bound [bit]
    DL_SR_WIDTH_MAX : UINT := 32;             // 位宽上限 [bit] / width upper bound [bit]
    DL_SR_LAST_BIT  : UINT := 31;             // 最高位号 [位] / the highest bit index [bit]
    DL_SR_CNT_MAX   : UDINT := 16#FFFF_FFFE;  // 计数饱和值 [次] / counter saturation value [times]
    DL_SR_MASK32    : DWORD := 16#FFFF_FFFF;  // 全宽掩码，宽度 32 时使用 [位图] / full width mask used at width 32 [bitmap]
    DL_SR_BIT31     : DWORD := 16#8000_0000;  // 最高位掩码，宽度 32 时提取溢出位 [位图] / top bit mask for the overflow extract at width 32 [bitmap]
    DL_SR_BIT0      : DWORD := 16#0001;       // 最低位掩码 [位图] / least significant bit mask [bitmap]
    DL_SR_ZERO      : DWORD := 16#0000;       // 零值常量，避免裸字面量 [位图] / zero constant, avoids a bare literal [bitmap]
    DL_SR_ONE       : DWORD := 16#0001;       // 一值常量，掩码减法用 [位图] / one constant used by the mask subtraction [bitmap]
    DL_SR_SHIFT_ONE : UINT := 1;              // 单步移位量与位宽步长 [bit] / single step shift amount and width step [bit]
END_VAR

// 段 1｜边沿实例无条件周期刷新（红线：严禁放入条件分支）/ segment 1, unconditional edge refresh
fbTrigShift(CLK := bShift);
fbTrigReset(CLK := bReset);

// 段 2｜输出与错误状态预置：脉冲量每拍先清 / segment 2, preset outputs and error status
bShiftOut := FALSE;                           // 单拍脉冲先清 / clear the single-cycle pulse first
bAnySet := FALSE;                             // 占位清零，段 7 重算 / clear, recomputed in segment 7
uSetCount := 0;                               // 置位计数先清 / clear the set-bit counter
eErr := 0;                                    // 预置无错误 / preset no error
bError := FALSE;                              // 预置无故障 / preset no fault

// 段 3｜使能闸：失能冻结寄存器，仅清脉冲 / segment 3, enable gate freezes the register
IF NOT bEnable THEN
    bAnySet := (uReg AND DL_SR_MASK32) <> DL_SR_ZERO; // 冻结态仍如实镜像非零判定 / still mirror the non-zero test while frozen
    RETURN;                                   // 失能即出口 / disabled is the exit
END_IF

// 段 4｜位宽闸：越界即故障级，寄存器清零且绝不索引任何位 / segment 4, width gate
IF (uWidth < DL_SR_WIDTH_MIN) OR (uWidth > DL_SR_WIDTH_MAX) THEN
    eErr := 16#0001_032A;                     // 位宽非法故障码 / illegal width fault id
    bError := TRUE;                           // 置故障标志 / raise the error flag
    uReg := DL_SR_ZERO;                       // 寄存器清零 / clear the register
    bShiftOut := FALSE;                       // 脉冲撤销 / drop the pulse
    bAnySet := FALSE;                         // 非零判定回 FALSE / non-zero test back to FALSE
    uSetCount := 0;                           // 置位计数回 0 / set-bit counter back to zero
    RETURN;                                   // 故障级提前返回，不触碰任何位 / early return, no bit is touched
END_IF

// 段 5｜掩码与移入位掩码构造（宽度 32 时走常量，禁 SHL(x, 32)）/ segment 5, mask construction
uWidthEff := uWidth;                          // 位宽已由段 4 保证在 1~32 / the width is guaranteed 1~32 by segment 4
IF uWidthEff >= DL_SR_WIDTH_MAX THEN
    uMask := DL_SR_MASK32;                    // 全宽掩码常量路径 / constant path for the full width
    uInMask := DL_SR_BIT31;                   // 最高位掩码常量路径 / constant path for the top bit
ELSE
    uMask := SHL(DL_SR_BIT0, uWidthEff) - DL_SR_ONE; // 2^n − 1，移位量 ≤ 31 结构性安全 / 2 to the n minus one, the shift never exceeds 31
    uInMask := SHL(DL_SR_BIT0, uWidthEff - DL_SR_SHIFT_ONE); // 最高有效位掩码，移位量 ≤ 31 / mask of the most significant effective bit
END_IF

// 段 6｜复位沿优先（清寄存器与计数）/ segment 6, reset edge has priority
IF fbTrigReset.Q THEN
    uReg := DL_SR_ZERO;                       // 寄存器清零 / clear the register
    uShiftCnt := 0;                           // 累计移位次数清零 / clear the accumulated shift count
END_IF

// 段 7｜清空优先于移位：安全侧宁可丢一位不可留脏位 / segment 7, clear has priority over shift
IF bClearAll THEN
    uReg := DL_SR_ZERO;                       // 整寄存器清零 / clear the whole register
    bShiftOut := FALSE;                       // 同拍不产生溢出位 / no overflow bit in the same cycle
    IF fbTrigShift.Q THEN
        eErr := 16#0001_0408;                 // 信息级：同拍清空与移位，已按清空优先 / info level, clearing wins in the same cycle
    END_IF
ELSIF fbTrigShift.Q THEN

    // 段 8｜提取溢出位（先取值再移位，顺序不可颠倒；溢出位跟随移位方向）/ segment 8, extract the overflow bit first, direction aware
    IF bDirLeft THEN
        bOutBit := (uReg AND uInMask) <> DL_SR_ZERO; // 左移：溢出位为最高有效位 / shifting left, the overflow bit is the most significant effective bit
    ELSE
        bOutBit := (uReg AND DL_SR_BIT0) <> DL_SR_ZERO; // 右移：溢出位为 bit0 / shifting right, the overflow bit is bit zero
    END_IF

    // 段 9｜移位并移入（移位量恒为 1，结构性小于位宽）/ segment 9, shift by one and insert
    IF bDirLeft THEN
        uReg := SHL(uReg, DL_SR_SHIFT_ONE);   // 向高位方向移一位，移位量 1 安全 / shift one position towards the higher bits
        IF bShiftIn THEN
            uReg := uReg OR DL_SR_BIT0;       // 低位端移入 / insert at the low end
        END_IF
    ELSE
        uReg := SHR(uReg, DL_SR_SHIFT_ONE);   // 向低位方向移一位 / shift one position towards the lower bits
        IF bShiftIn THEN
            uReg := uReg OR uInMask;          // 高位端移入 / insert at the high end
        END_IF
    END_IF

    // 段 10｜超宽截断：旧位残留在高位会造成假置位 / segment 10, truncate to the effective width
    uReg := uReg AND uMask;                   // 与有效掩码相与 / and with the effective mask
    bShiftOut := bOutBit;                     // 发布本拍溢出位 / publish the overflow bit

    // 段 11｜移位计数饱和（饱和即置码，绝不回绕）/ segment 11, saturating shift counter
    IF uShiftCnt < DL_SR_CNT_MAX THEN
        uShiftCnt := uShiftCnt + 1;           // 饱和加一 / saturating increment
    ELSE
        eErr := 16#0001_032B;                 // 故障级：统计量已不可信 / fault level, the statistics are no longer trustworthy
        bError := TRUE;                       // 置故障标志 / raise the error flag
    END_IF
END_IF

// 段 12｜置位统计（位宽已保证 ≤ 32，移位量 ≤ 31）/ segment 12, set-bit statistics
FOR uIdx := 0 TO uWidthEff - DL_SR_SHIFT_ONE DO
    IF (uReg AND SHL(DL_SR_BIT0, uIdx)) <> DL_SR_ZERO THEN
        uSetCount := uSetCount + 1;           // 逐位累加置位数 / accumulate the set bits one by one
    END_IF
END_FOR
bAnySet := uSetCount > 0;                     // 非零判定由计数导出，避免二次遍历 / derived from the count, no second pass
END_FUNCTION_BLOCK

(* ---- FB_DL_BlinkOutput.st ---- *)
(*
    FB_DL_BlinkOutput —— 方波闪烁输出（tOn / tOff 独立交替两相 TON）
    ------------------------------------------------------------------
    组件名称  : FB_DL_BlinkOutput
    分类      : DL_Base / SignalGeneration
    前缀      : FB_DL_
    版本      : 1.0.0
    溯源      : 借鉴组织 —— T1-1 OSCAT Basic（矩阵行 170）：仅借鉴 BLINK 的
                **公开行为定义**（tOn / tOff 独立交替两相 + 使能撤除冻结输出
                与相位），OSCAT 许可免费、按 EPL-2.0 类比先例（R25）致谢；
                clean-room 声明 —— **零代码行复制**，实现 / 引脚名 / 码位 /
                组态锁存口径 100% 自有。
    平台      : 纯 IEC 61131-3（双 TON 交替），CODESYS 3.5 / TwinCAT 3 /
                InoProShop / Machine Expert 通用
    作者      : 道莅代码库 · PLC编程专家（R72 构建轮 · 批 3 · 序号 8）
    ------------------------------------------------------------------
    功能说明  : 秒级方波闪烁：tOn 相（bOut = TRUE）计时满 tOn → 切 tOff 相
                （bOut = FALSE）→ 计满 tOff 回切开相，如此交替。真实工况：
                塔灯辅闪、报警闪烁、待机呼吸灯。
                相机制（两相判据链，无顺序状态机 CASE）：
                ① 双 TON 实例按当前相择一计时，IN 为显式条件变量；
                ② bEn = FALSE 冻结 bOut 与相位**计数值**（失能不清相位，恢复
                   时从冻结点续走——相位保持，定时清零重启，OSCAT BLINK 行为
                   定义口径）；失能期间双 TON 的 IN 强制 FALSE（计时同步冻结），
                   R191 失能语义声明：**冻结保持末值**（bOut 不清零）；
                ③ tOn = 0 或 tOff = 0（TIME 无负值路径）→ **组态锁存码**
                   （防全灭 / 全亮静默——fGain = 0 报警静默教训 R386 同型），
                   锁存至 bReset 上升沿唯一解除（R188，解除路径恒可达自证）；
                   锁存相 bOut 强制 FALSE、周期计数冻结（故障可见性靠码位 +
                   bError，不靠灯）；
                ④ 周期计数口径：每完成一个完整 on + off 周期（关相计满回切
                   开相瞬间）uCycleCount + 1，UDINT 饱和上限 16#FFFF_FFFF。
                段序口径：锁存（含解除与首次成因登记）先于定时器调用——
                消灭「零组态拍定时器先跑一拍」的伪切换伪影；双 TON 与
                R_TRIG 仍为每拍无条件调用（IN 显式条件，选相不进可跳过分支）。
                TON 极性声明（R319 复核）：双 TON 的 IN = 相内剩余条件
                （_bRun AND 相标志），**非**被监视正常电平——本件是相驱动
                而非监视件，极性合规。
    错误码    : 16#0001_0752 组态非法：tOn = 0 或 tOff = 0（零时长相会退化
                            为全灭或全亮静默），锁存至复位沿 —— 故障级
                加码反证句（R90）：该场景无法由「正常闪烁输出 + bValid」
                观测——正常相 bOut 在闪烁、锁存相 bOut 恒 FALSE + bError =
                TRUE + 码位回放，输出组合不可互换，故立独立码。
    码位总账  : 16#0001_0752 用（同段 16#0001_0753 已由 FC_DL_DaysInMonthChk
                占用，本件不占）
    状态机    : 无顺序状态机 CASE——两相判据链 + 双 TON 自持；非法状态不可能
                出现（_bPhaseOn 为 BOOL，无非法值域）
    边界与披露: 一 双 TON（tonOn / tonOff）与 R_TRIG（rtReset）每拍
                   **无条件调用**（规则 ⑦），IN 为显式条件变量；
                二 零全局变量、零 VAR_EXTERNAL、零物理地址；
                三 组态域闸逐项点名（R272）：tOn / tOff 双引脚全部纳入零值
                   锁存闸；
                四 验收向量：tOn = tOff 恰等（对称方波）→ 正常 50% 占空比；
                   tOn / tOff 极端幅值 T#1E9MS（约 11.6 天）→ 正常慢闪
                   （TIME 32 位 ms 域内可表，无溢出面）；tOn = T#0MS →
                   0752 锁存；V5 失能 → bOut 冻结、相位保持、计数冻结；
                   V6 复位沿解除锁存后恢复闪烁；
                五 同拍双窗配比约束（R100）：双相独立计时无窗间依赖约束
                （tOn / tOff 各自独立，无先后门槛），配比约束句豁免声明；
                六 输出语义：uCycleCount 饱和口径（16#FFFF_FFFF 封顶不再
                   累加，防回绕）；
                七 依赖声明：仅 Standard.library（TON / R_TRIG），零厂商方言。
    验收向量  : V1 tOn = T#1S，tOff = T#1S → 50% 对称方波；
                V2 tOn = T#0MS → 0752 锁存 + bError；V3 tOff = T#0MS →
                0752 锁存；V4 tOn = T#500MS，tOff = T#2S → 20% 占空比；
                V5 bEn 置 FALSE → bOut 与 _bPhaseOn 冻结；V6 bReset 上升沿
                → 解锁恢复；V7 一个完整周期后 uCycleCount = 1。
                算法已证（脚本）：未跑 ｜ 编译器已证（三平台）：未跑
    修订记录  : 2026-11-23 v1.0.0 首次入库（R72 构建轮 · 批 3 · 序号 8）
*)
FUNCTION_BLOCK FB_DL_BlinkOutput
VAR_INPUT
    bEn    : BOOL := FALSE;                (* 使能，[标志]，FALSE 冻结输出与相位（R191 冻结保持声明）/ the enable, FALSE freezes the output and the phase *)
    tOn    : TIME := T#500MS;              (* 开相时长，[ms]，禁 0（零值锁存 0752）/ the on phase duration, must not be zero *)
    tOff   : TIME := T#500MS;              (* 关相时长，[ms]，禁 0（零值锁存 0752）/ the off phase duration, must not be zero *)
    bReset : BOOL := FALSE;                (* 组态故障复位，[标志]，上升沿唯一解除（R188）/ the configuration fault reset, its rising edge is the only release *)
END_VAR
VAR_OUTPUT
    bOut        : BOOL := FALSE;           (* 方波输出，[标志]，失能冻结保持末值 / the square wave output, frozen on disable *)
    uCycleCount : UDINT := 0;              (* 完整周期计数（on + off 计满一回切加一），饱和上限 16#FFFF_FFFF [次] / the complete cycle count, saturated *)
    bValid      : BOOL := FALSE;           (* 出口可用标志，锁存故障为 FALSE / the outlets usable flag *)
    bError      : BOOL := FALSE;           (* 故障标志，与锁存同源（R191）/ the fault flag from the latch *)
    nErrCode    : UDINT := 16#0000_0000;   (* 错误码，0 = 正常，锁存回放（R187）/ the error id, replayed from the latch *)
END_VAR
VAR
    _bPhaseOn  : BOOL := TRUE;             (* 相位寄存器：TRUE = 开相（上电首拍从开相起走）/ the phase register, TRUE for the on phase *)
    _bFault    : BOOL := FALSE;            (* 组态故障锁存副本，仅复位沿解除 / the config fault latch copy *)
    _nCodeLatch: UDINT := 0;               (* 锁存成因码，故障期回放 / the latched cause code *)
    _bRun      : BOOL := FALSE;            (* 运行许可 = 使能 且 无锁存故障 / the run permit *)
    tonOn      : TON;                      (* 开相计时实例，每拍无条件调用 / the on phase timer *)
    tonOff     : TON;                      (* 关相计时实例，每拍无条件调用 / the off phase timer *)
    rtReset    : R_TRIG;                   (* 复位沿实例，每拍无条件调用 / the reset edge instance *)
END_VAR
VAR CONSTANT
    DL_BLO_TZERO  : TIME := T#0S;          (* 零时长哨兵（组态锁存闸）[ms] / the zero duration sentinel *)
    DL_BLO_CYCMAX : UDINT := 16#FFFF_FFFF; (* 周期计数饱和上限 [次] / the cycle count saturation cap *)
    DL_BLO_CODE   : UDINT := 16#0001_0752; (* 组态非法锁存码 [码] / the illegal configuration latch code *)
    DL_BLO_ZERO   : UDINT := 0;            (* 无符号零哨兵 [码] / the unsigned zero sentinel *)
    DL_BLO_ONE    : UDINT := 1;            (* 计数步进 [次] / the count step *)
END_VAR

// 段 0｜复位沿无条件调用（规则 ⑦）/ segment 0, the unconditional reset edge refresh
rtReset(CLK := bReset);                    // 每拍无条件刷新 / refreshed every scan without exception

// 段 1｜锁存解除与首次成因登记（先锁存后计时，消灭零组态拍伪切换伪影）/ segment 1, the latch release and the first cause registration
IF rtReset.Q THEN                          // 复位上升沿 / the reset rising edge
    _bFault := FALSE;                      // 解除锁存（唯一解除边，R188，恒可达 R152 自证）/ release the latch
    _nCodeLatch := DL_BLO_ZERO;            // 清锁存码（作用域声明 R311：仅清锁存与码，不清相位与计数）/ clear the latched code
END_IF
IF (NOT _bFault) AND ((tOn = DL_BLO_TZERO) OR (tOff = DL_BLO_TZERO)) THEN // 零时长相组态命中 / a zero duration configuration hit
    _bFault := TRUE;                       // 置锁存（防全灭 / 全亮静默，R386 同型）/ latch the fault
    _nCodeLatch := DL_BLO_CODE;            // 登记成因码（首次成因锁存，故障期不重推断 R189）/ register the cause code
END_IF

// 段 2｜运行许可与双 TON 无条件调用（IN 为显式条件变量，选相不进可跳过分支）/ segment 2, the run permit and the unconditional timer calls
_bRun := bEn AND (NOT _bFault);            // 运行许可（锁存已定，无伪影）/ the run permit
tonOn(IN := _bRun AND _bPhaseOn, PT := tOn);         // 开相计时（失能 / 关相时 IN FALSE 冻结）/ the on timer
tonOff(IN := _bRun AND (NOT _bPhaseOn), PT := tOff); // 关相计时 / the off timer

// 段 3｜两相交替推进（运行许可内；失能 / 故障相不动相位与计数）/ segment 3, the two phase progression
IF _bRun THEN                              // 运行许可成立 / the run permit holds
    IF _bPhaseOn THEN                      // 开相 / the on phase
        bOut := TRUE;                      // 输出亮 / the output on
        IF tonOn.Q THEN                    // 开相计满 / the on phase timed out
            _bPhaseOn := FALSE;            // 切关相 / switch to the off phase
        END_IF
    ELSE                                   // 关相 / the off phase
        bOut := FALSE;                     // 输出灭 / the output off
        IF tonOff.Q THEN                   // 关相计满（完整 on + off 周期完成）/ the off phase timed out
            _bPhaseOn := TRUE;             // 回切开相 / back to the on phase
            IF uCycleCount < DL_BLO_CYCMAX THEN // 饱和上限闸（防回绕）/ the saturation cap
                uCycleCount := uCycleCount + DL_BLO_ONE; // 周期计数 + 1 / count one cycle
            END_IF
        END_IF
    END_IF
ELSIF _bFault THEN                         // 锁存故障相（故障可见性靠码位与 bError）/ the latched fault phase
    bOut := FALSE;                         // 故障相强制灭（不冻结残留亮态）/ force off in the fault phase
END_IF                                     // 失能相（非故障）：bOut 不触碰，冻结保持（R191 声明）

// 段 4｜统一出口（名实双出口同源，R191）/ segment 4, the unified outlet
bValid := NOT _bFault;                     // 出口可用 = 无锁存 / the usable flag
bError := _bFault;                         // 故障标志与锁存同源 / the flag shares the latch
IF _bFault THEN                            // 锁存回放（R187）/ the latched replay
    nErrCode := _nCodeLatch;               // 回放锁存码 / replay the latched code
ELSE                                       // 正常相 / the normal phase
    nErrCode := DL_BLO_ZERO;               // 无错 / ok
END_IF
END_FUNCTION_BLOCK

(* ---- FB_DL_ClockDriftMonitor.st ---- *)
(*==============================================================================
 * 组件名称 (Component)  : FB_DL_ClockDriftMonitor
 * 所属子库 (Sublibrary) : DL_Base
 * 当前版本 (Version)    : 1.0.1
 * 兼容性   (Platform)   : CODESYS 3.5 / TwinCAT 3 / 汇川 InoProShop / Machine Expert
 *                         仅依赖 Standard.library（TON / R_TRIG / SUB / TIME_TO_REAL），
 *                         SUB(DT,DT)->TIME 为 IEC 61131-3 标准函数表语义，零厂商方言
 * 来源标签 (Source)     : self-std
 * 功能描述 (Function)   : 本地 RTC 对外部标准钟的漂移率监视：每个采样窗分别求两钟
 *                         相对上一窗基线的时间增量，差值即窗内漂移量 [ms]，折算为
 *                         漂移率 [ms/h]（LREAL 承载防溢出），经 5 样本滑动窗中位滤波
 *                         后与漂移率上限比较产生告警；累计漂移超同步阈值置「需校钟」。
 *                         钟回拨（任一钟相对上窗基线负跳）单列「校钟事件」：只置事件
 *                         不计漂移、不置告警，并就地重立基线。
 *                         本件只监视不写钟——写钟归系统层，本件零输出侧钟操作。
 * 边界与语义披露 (Boundary disclosure) :
 *   1) 两钟均以 DT 引脚注入（零全局耦合）；DT 零值（DT#1970-01-01-00:00:00）视为
 *      未初始化，按故障级锁存，两钟各自独立码位（归因唯一 R190）。
 *   2) 窗增量以 TIME 承载：两钟相邻窗基线间隔超过 IEC TIME 正域上限（约 24.8 天，
 *      有符号口径）时增量回绕为巨值——以 3.0E9 ms（约 34.7 天）界作回绕哨兵，
 *      触发按「校钟事件」处理并重立基线，绝不把回绕值折算成漂移率。
 *   3) 首窗只立基线不发布漂移（无前窗可比），基线窗与运行窗状态分离。
 *   4) 漂移率与累计漂移的正负号语义：正 = 本地钟慢于外部标准钟（本地增量不足），
 *      负 = 本地钟快；告警与需校钟判据均取绝对值。
 *   5) SUB(DT,DT) 与 DT 比较（<）均为 IEC 61131-3 标准函数/运算语义。
 *      交付门槛：须在 CODESYS / TwinCAT / InoProShop 三平台各编译验证一次（R64）。
 * 故障码表 (Error codes) :
 *   16#0001_03EF [故障级] 外部标准钟无效（DT 零值未初始化），锁存至复位沿
 *                 反证：该场景下漂移率恒不发布（fDriftRateMsH 保持末值）、
 *                 状态 eFault——但 eFault 无法区分是哪只钟无效，需独立码位。
 *   16#0001_03F0 [故障级] 本地 RTC 无效（DT 零值未初始化），锁存至复位沿
 *                 反证：本地钟失效与外部钟失效对 eState / 漂移不发布等输出的影响组合完全一致，不可区分。
 *   16#0001_03F1 [故障级] 采样窗组态非法（<= T#0S），拒绝采样，锁存至复位沿
 *                 反证：窗非法时无窗脉冲（bWindowTick 恒 FALSE）与「使能关闭」
 *                 输出组合相同，无码不可区分。
 *   16#0001_04B3 [信息级] 中位滤波后漂移率超限（告警确认）
 *                 反证：bDriftAlarm 已是保持型位，但超限方向（快/慢）不可由
 *                 布尔位观测，码位承载「已确认超限」事实供 HMI 记录。
 *   16#0001_04B4 [信息级] 钟回拨 / 窗增量回绕，已按校钟事件重立基线
 *                 反证：回拨拍 bSyncEvent 为单拍脉冲，事件落账后即消失，
 *                 无码则历史回拨次数不可考。
 *   16#0001_04B5 [信息级] 累计漂移超同步阈值（需校钟确认）
 *                 反证：bNeedSync 为保持型位，码位用于事件流水归档，与告警码
 *                 分开承载两类不同事实（率超限 vs 累计超限）。
 *   非法状态拦截复用全库惯用码 16#0001_0005（不新占号）。
 * 码位总账 (Code ledger) : 16#0001_03EF / 03F0 / 03F1 用 ｜ 16#0001_04B3 / 04B4 / 04B5 用
 * 依赖     (Depends)    : 无 DL_ 内部依赖；Standard.library: TON / R_TRIG / SUB / TIME_TO_REAL
 * 红线自检 (Redline)    : R1 ✓ 零全局变量与 VAR_EXTERNAL ｜ R2 ✓ 零 %I/%Q 物理地址
 *                         R3 ✓ 纯 IEC 61131-3（SUB/TIME_TO_REAL 均标准语义）
 *                         R4 ✓ 窗判零 / 折算分母 eps 闸 / 非有限双判（自反 + 差自减）
 *                         R5 ✓ 全变量中英双语同行注释 ｜ R6 ✓ 四态 ENUM + CASE + ELSE 兜底
 *                         R7 ✓ 二沿一计时主体最前部无条件刷新；窗 TON 自复位（IN 串自身 Q 取反）
 * 修订历史 (Revision)   :
 *   2026-11-22  v1.0.0  首版入库（R68 构建轮 · 批 1 · 目标 2）
 *   2026-11-22  v1.0.1  终审就地修①：组态锁存解除路径可达化（复位沿 + 三类非法源消失即清锁存，原 eFault 相不可达）
 *============================================================================*)

(*-----------------------------------------------------------------------------
 * 枚举: E_DL_ClockDriftState（归属 DL_Base，与 FB_DL_ClockDriftMonitor 同文件）
 *----------------------------------------------------------------------------*)
TYPE E_DL_ClockDriftState :
(
    eIdle     := 0,    // 未使能：全部告警与累计量冻结 / Disabled, alerts and accumulators frozen
    eBaseline := 10,   // 等待首窗基线：只存钟不发布 / Awaiting first window baseline, no publish
    eRun      := 20,   // 采样运行：每窗发布漂移率 / Running, drift rate published per window
    eFault    := 99    // 组态 / 钟源无效锁存 / Config or clock source latched invalid
);
END_TYPE

(*==============================================================================
 * 功能块: FB_DL_ClockDriftMonitor
 * 调用约定: 每个扫描周期无条件调用一次；两钟 DT 引脚须每拍刷新注入。
 *============================================================================*)
FUNCTION_BLOCK FB_DL_ClockDriftMonitor
VAR_INPUT
    dtExtStd         : DT;                     // 外部标准钟快照 [UTC]，零值 = 未初始化 / External standard clock, zero = uninitialized
    dtLocRtc         : DT;                     // 本地 RTC 快照 [本地]，零值 = 未初始化 / Local RTC snapshot, zero = uninitialized
    tSampleWin       : TIME  := T#30M;         // 采样窗时长 [min]，<= T#0S 组态非法 / Sampling window [min], <= 0 illegal
    fRateLimitMsH    : LREAL := 100.0;         // 漂移率告警上限 [ms/h] / Drift rate alarm limit [ms per hour]
    fSyncThresholdMs : LREAL := 5000.0;        // 累计漂移需校钟阈值 [ms] / Cumulative drift sync threshold [ms]
    bEnable          : BOOL  := TRUE;          // 监视使能 / Monitor enable
    bAckSync         : BOOL;                   // 上升沿：校钟完成确认，清累计漂移 / Rising edge: sync done, clears cumulative drift
    bReset           : BOOL;                   // 上升沿：清除钟源 / 组态故障锁存 / Rising edge: clears source and config latches
END_VAR
VAR_OUTPUT
    fDriftRateMsH : LREAL;                   // 中位滤波后漂移率 [ms/h] / Median filtered drift rate [ms per hour]
    fDriftRawMsH  : LREAL;                   // 本窗原始漂移率 [ms/h]，诊断 / Raw drift rate of the last window
    fCumDriftMs   : LREAL;                   // 累计漂移 [ms]，正 = 本地慢 / Cumulative drift [ms], positive = local slow
    bDriftAlarm   : BOOL;                    // 漂移率超限告警（保持型）/ Drift rate over limit alarm, level held
    bNeedSync     : BOOL;                    // 需校钟（累计超阈值，保持型）/ Sync required, level held
    bSyncEvent    : BOOL;                    // 校钟事件脉冲（回拨 / 回绕，单拍）/ Sync event pulse, single scan
    bWindowTick   : BOOL;                    // 采样窗脉冲（单拍，诊断）/ Window tick pulse, single scan, diagnostics
    bError        : BOOL;                    // 故障标志（钟源 / 组态锁存）/ Fault flag, source or config latched
    uErrorId      : UDINT;                   // 故障码，0 = 无故障 / Error code, 0 = none
    eState        : E_DL_ClockDriftState;    // 当前状态（供 HMI 诊断）/ Current state for HMI diagnosis
END_VAR
VAR
    fbTrigAck     : R_TRIG;                  // 校钟确认沿检测实例 / Sync acknowledge edge detector
    fbTrigReset   : R_TRIG;                  // 复位沿检测实例 / Reset edge detector
    tonWin        : TON;                     // 采样窗计时（自复位）实例 / Sampling window timer, self resetting
    eStateInt     : E_DL_ClockDriftState;    // 主状态机内部当前态 / Internal state machine state
    dtExtPrev     : DT;                      // 上窗外部标准钟基线 / Previous window external baseline
    dtLocPrev     : DT;                      // 上窗本地钟基线 / Previous window local baseline
    tDeltaExt     : TIME;                    // 本窗外部钟增量 [ms] / External clock delta this window [ms]
    tDeltaLoc     : TIME;                    // 本窗本地钟增量 [ms] / Local clock delta this window [ms]
    fMsExt        : LREAL;                   // 外部钟增量实数化 [ms] / External delta as LREAL [ms]
    fMsLoc        : LREAL;                   // 本地钟增量实数化 [ms] / Local delta as LREAL [ms]
    fDriftMs      : LREAL;                   // 本窗漂移量 [ms] / Drift amount this window [ms]
    fWinHours     : LREAL;                   // 窗长折算小时 [h] / Window length in hours [h]
    fRateRaw      : LREAL;                   // 原始漂移率中间量 [ms/h] / Raw drift rate intermediate
    afRateRing    : ARRAY[0..4] OF LREAL;    // 漂移率滑动窗 [ms/h]，5 样本 / Drift rate sliding window, 5 samples
    afRateSort    : ARRAY[0..4] OF LREAL;    // 中位排序暂存区 / Median sort scratch
    nRingWrite    : INT;                     // 滑动窗写指针 [0..4] / Sliding window write pointer
    nRingFill     : INT;                     // 滑动窗已填样本数 [个] / Filled sample count
    nI            : INT;                     // 排序外层索引 / Sort outer index
    nJ            : INT;                     // 排序内层索引 / Sort inner index
    fKey          : LREAL;                   // 插入排序当前键值 / Insertion sort key
    fCumInt       : LREAL;                   // 累计漂移内部副本 [ms] / Internal cumulative drift [ms]
    bExtInvalid   : BOOL;                    // 本拍外部钟无效 / External clock invalid this scan
    bLocInvalid   : BOOL;                    // 本拍本地钟无效 / Local clock invalid this scan
    bWinInvalid   : BOOL;                    // 本拍采样窗组态非法 / Window config illegal this scan
    bFaultLatch   : BOOL;                    // 故障锁存（复位沿清除）/ Fault latch, cleared by reset edge
    bErrorInt     : BOOL;                    // 本拍故障置位累加（出口归并）/ Fault set accumulator of this scan
    bFirstScan    : BOOL := TRUE;            // 上电首扫标志 / First-scan flag
END_VAR
VAR CONSTANT
    DL_CD_RING_CAP  : INT   := 5;            // 中位滤波窗容量 [个] / Median window capacity
    DL_CD_MEDIAN_MID: INT   := 2;            // 5 样本中位下标 / Median index of 5 samples
    DL_CD_WRAP_MS   : LREAL := 3.0E9;        // 窗增量回绕哨兵 [ms]，约 34.7 天 / Window delta wrap sentinel [ms]
    DL_CD_HOUR_MS   : LREAL := 3600000.0;    // 小时毫秒换算常数 [ms/h] / Hours to milliseconds factor
    DL_CD_EPS       : LREAL := 1.0E-9;       // 窗长折算判零容差 [h] / Window length zero tolerance [h]
    DL_CD_CUM_MAX   : LREAL := 1.0E12;       // 累计漂移饱和上限 [ms] / Cumulative drift saturation [ms]
END_VAR

(*------------------------------------------------------------------------------
 * 段 1｜无条件刷新区（红线 R7）：二沿 + 窗计时（IN 串 bEnable AND NOT 自身 Q，自复位 R188）
 *      Unconditional refresh: two edges plus the self resetting window timer
 *-----------------------------------------------------------------------------*)
fbTrigAck(CLK := bAckSync);
fbTrigReset(CLK := bReset);
tonWin(IN := bEnable AND (NOT tonWin.Q), PT := tSampleWin);

(*------------------------------------------------------------------------------
 * 段 2｜上电首扫：基线钟显式落零哨兵（与零值 = 未初始化闸共用判据，不误发故障）
 *      First-scan init: baselines forced to the zero sentinel, sharing the gate
 *-----------------------------------------------------------------------------*)
IF bFirstScan THEN
    dtExtPrev  := dtExtStd;
    dtLocPrev  := dtLocRtc;
    eStateInt  := E_DL_ClockDriftState.eBaseline;
    nRingWrite := 0;
    nRingFill  := 0;
    fCumInt    := 0.0;
    bFirstScan := FALSE;
END_IF

(*------------------------------------------------------------------------------
 * 段 3｜每拍预清（FB32-1）：单拍位统一预置，禁入锁存 / 快照 / 累计量
 *      Per-scan preset: single-scan flags only
 *-----------------------------------------------------------------------------*)
bErrorInt   := FALSE;
bSyncEvent  := FALSE;
bWindowTick := FALSE;

(*------------------------------------------------------------------------------
 * 段 4｜组态域闸（R151 / R190 归因唯一）：两钟零值各自独立码位 + 窗判零
 *      Config gate: each clock gets its own code, plus the window zero gate
 *      DT 与 DT#1970-01-01-00:00:00 精确相等比较（离散类型直比合法，非浮点）
 *-----------------------------------------------------------------------------*)
bExtInvalid := (dtExtStd = DT#1970-01-01-00:00:00);
bLocInvalid := (dtLocRtc = DT#1970-01-01-00:00:00);
bWinInvalid := (tSampleWin <= T#0S);

IF bExtInvalid OR bLocInvalid OR bWinInvalid THEN
    bFaultLatch := TRUE;
END_IF

(* 终审就地修 v1.0.1（R68）：解除路径（R152 自证可达）——复位沿 AND 组态非法条件
 * 全部消失即清锁存。原实现把锁存清零只写在 eFault 相分支，而组态闸置锁存后
 * 并不迁相至 eFault（只回 eIdle / 驻留），eFault 相不可达 -> 锁存永不可解，
 * 组件保护/监视功能一次性永久失效直至 PLC 重启（终审两式①）。
 * Clear path made provably reachable: reset edge with the illegal config gone. *)
IF fbTrigReset.Q AND (NOT bExtInvalid) AND (NOT bLocInvalid) AND (NOT bWinInvalid) THEN
    bFaultLatch := FALSE;         // 锁存解除 / Latch cleared
    uErrorId    := 16#0000_0000;  // 码位随解除归零 / Code cleared with the latch
END_IF

IF bExtInvalid THEN
    uErrorId  := 16#0001_03EF;    // 故障级：外部标准钟无效 / Fault: external clock invalid
    bErrorInt := TRUE;
ELSIF bLocInvalid THEN
    uErrorId  := 16#0001_03F0;    // 故障级：本地 RTC 无效 / Fault: local RTC invalid
    bErrorInt := TRUE;
ELSIF bWinInvalid THEN
    uErrorId  := 16#0001_03F1;    // 故障级：采样窗组态非法 / Fault: window config illegal
    bErrorInt := TRUE;
END_IF

(*------------------------------------------------------------------------------
 * 段 5｜校钟确认沿：清累计漂移（作用域声明：只清累计量，不清基线与告警）
 *      Sync acknowledge edge: clears the cumulative drift only
 *-----------------------------------------------------------------------------*)
IF fbTrigAck.Q THEN
    fCumInt := 0.0;               // 累计漂移归零（作用域：仅累计量）/ Clear cumulative only
END_IF

(*------------------------------------------------------------------------------
 * 段 6｜主状态机（红线 R6）：ENUM + CASE + ELSE 兜底
 *      Main state machine with the mandatory ELSE fallback
 *-----------------------------------------------------------------------------*)
CASE eStateInt OF

    E_DL_ClockDriftState.eIdle:
        IF bEnable AND (NOT bFaultLatch) THEN
            dtExtPrev := dtExtStd;     // 重入先立新基线 / New baseline on re-entry
            dtLocPrev := dtLocRtc;
            eStateInt := E_DL_ClockDriftState.eBaseline;
        END_IF

    E_DL_ClockDriftState.eBaseline:
        (* eWait 类相退出条件 >= 2 条（R98）：窗脉冲沿 + 进相前置消失（失能 / 故障） *)
        IF bFaultLatch OR (NOT bEnable) THEN
            eStateInt := E_DL_ClockDriftState.eIdle;
        ELSIF tonWin.Q THEN
            dtExtPrev := dtExtStd;     // 首窗只立基线不发布 / First window stores baseline only
            dtLocPrev := dtLocRtc;
            eStateInt := E_DL_ClockDriftState.eRun;
        END_IF

    E_DL_ClockDriftState.eRun:
        IF bFaultLatch OR (NOT bEnable) THEN
            eStateInt := E_DL_ClockDriftState.eIdle;
        ELSIF tonWin.Q THEN
            bWindowTick := TRUE;       // 窗脉冲（诊断）/ Window tick for diagnostics
            IF (dtLocRtc < dtLocPrev) OR (dtExtStd < dtExtPrev) THEN
                (* 回拨（差值负跳）：只置校钟事件不计漂移不置告警，就地重立基线 *)
                (* Rollback: sync event only, no drift, no alarm, re-baseline *)
                bSyncEvent := TRUE;
                uErrorId   := 16#0001_04B4;
                dtExtPrev  := dtExtStd;
                dtLocPrev  := dtLocRtc;
            ELSE
                tDeltaExt := SUB(dtExtStd, dtExtPrev);   // 外部钟窗增量 / External window delta
                tDeltaLoc := SUB(dtLocRtc, dtLocPrev);   // 本地钟窗增量 / Local window delta
                fMsExt := TIME_TO_LREAL(tDeltaExt);
                fMsLoc := TIME_TO_LREAL(tDeltaLoc);
                IF (fMsExt >= DL_CD_WRAP_MS) OR (fMsLoc >= DL_CD_WRAP_MS) THEN
                    (* 窗增量回绕哨兵触发：按校钟事件处理，绝不折算漂移率 *)
                    (* Wrap sentinel hit: treated as a sync event, never scaled *)
                    bSyncEvent := TRUE;
                    uErrorId   := 16#0001_04B4;
                ELSE
                    fDriftMs  := fMsExt - fMsLoc;        // 窗内漂移量 [ms] / Window drift [ms]
                    fWinHours := TIME_TO_LREAL(tSampleWin) / DL_CD_HOUR_MS;
                    IF fWinHours > DL_CD_EPS THEN
                        fRateRaw := fDriftMs / fWinHours;  // 折算漂移率 [ms/h]，分母已闸 / Rate, guarded denominator
                        IF (fRateRaw <> fRateRaw) OR ((fRateRaw - fRateRaw) <> (fRateRaw - fRateRaw)) THEN
                            (* 非有限兜底三件套（R258）：冻结发布 + 故障码 + bError + 不发布 *)
                            fRateRaw  := 0.0;
                            uErrorId  := 16#0001_0005;
                            bErrorInt := TRUE;
                        ELSE
                            fDriftRawMsH := fRateRaw;
                            fDriftRateMsH := MedianOfRing(fRateRaw);  // 中位滤波委托 / Median via private method
                            IF ABS(fDriftRateMsH) > fRateLimitMsH THEN
                                bDriftAlarm := TRUE;           // 告警置位（保持型）/ Level alarm set
                                uErrorId    := 16#0001_04B3;   // 信息级：率超限确认 / Info: rate confirmed
                            ELSIF ABS(fDriftRateMsH) <= fRateLimitMsH THEN
                                bDriftAlarm := FALSE;          // 回落清除（与阈值同点，无回差）/ Clear on recovery
                            END_IF
                            IF ABS(fCumInt) < DL_CD_CUM_MAX THEN
                                fCumInt := fCumInt + fDriftMs; // 累计推进（饱和守卫）/ Accumulate, guarded
                            END_IF
                            IF ABS(fCumInt) > fSyncThresholdMs THEN
                                bNeedSync := TRUE;             // 需校钟置位 / Sync required set
                                uErrorId  := 16#0001_04B5;     // 信息级：累计超限确认 / Info: cumulative confirmed
                            ELSE
                                bNeedSync := FALSE;            // 确认沿已归零后回落清除 / Clear after ack
                            END_IF
                        END_IF
                    END_IF
                END_IF
                dtExtPrev := dtExtStd;     // 窗尾统一刷新基线 / Baselines refreshed at window tail
                dtLocPrev := dtLocRtc;
            END_IF
        END_IF

    E_DL_ClockDriftState.eFault:
        (* 解除路径（R152 自证可达）：复位沿 AND 三类非法源全部消失 *)
        IF fbTrigReset.Q AND (NOT bExtInvalid) AND (NOT bLocInvalid) AND (NOT bWinInvalid) THEN
            bFaultLatch := FALSE;
            bDriftAlarm := FALSE;
            bNeedSync   := FALSE;
            uErrorId    := 16#0000_0000;
            eStateInt   := E_DL_ClockDriftState.eIdle;
        END_IF

    ELSE
        (* 非法状态拦截：不做隐式恢复，直接锁存上报 *)
        eStateInt := E_DL_ClockDriftState.eFault;
        uErrorId  := 16#0001_0005;
        bErrorInt := TRUE;

END_CASE;

(*------------------------------------------------------------------------------
 * 段 7｜输出单一出口（范式 P-05）
 *      Single output exit
 *-----------------------------------------------------------------------------*)
fCumDriftMs := fCumInt;
bError := bErrorInt OR (eStateInt = E_DL_ClockDriftState.eFault);
eState := eStateInt;
END_FUNCTION_BLOCK

(*------------------------------------------------------------------------------
 * 私有方法: MedianOfRing —— 滑动窗写入 + 插入排序取中位（5 样本固定容量，无死循环风险）
 *      Private method: ring write plus insertion sort median over 5 fixed slots
 *      调用约定: 仅在 eRun 相窗脉冲拍调用；两层循环边界均为常量，开闭词配对
 *----------------------------------------------------------------------------*)
METHOD MedianOfRing : LREAL
VAR_INPUT
    fNew : LREAL;    // 本窗新样本 [ms/h] / New sample of this window [ms per hour]
END_VAR

afRateRing[nRingWrite] := fNew;                       // 新样本入环 / New sample into the ring
nRingWrite := nRingWrite + 1;
IF nRingWrite >= DL_CD_RING_CAP THEN
    nRingWrite := 0;                                  // 显式回卷 / Explicit wrap
END_IF
IF nRingFill < DL_CD_RING_CAP THEN
    nRingFill := nRingFill + 1;                       // 填充计数推进 / Fill count up
END_IF

IF nRingFill < 3 THEN
    MedianOfRing := fNew;    // 样本不足 3 个：中位未定义，直通新样本（R307 挂起语义）/ Fewer than 3 samples: pass through
    RETURN;
END_IF

FOR nI := 0 TO (nRingFill - 1) DO                     // 复制有效区到排序暂存 / Copy valid span
    afRateSort[nI] := afRateRing[nI];
END_FOR

FOR nI := 1 TO (nRingFill - 1) DO                     // 插入排序（升序）/ Insertion sort ascending
    fKey := afRateSort[nI];
    nJ  := nI - 1;
    WHILE (nJ >= 0) AND (afRateSort[nJ] > fKey) DO    // 内层右移 / Inner shift right
        afRateSort[nJ + 1] := afRateSort[nJ];
        nJ := nJ - 1;
    END_WHILE
    afRateSort[nJ + 1] := fKey;
END_FOR

MedianOfRing := afRateSort[DL_CD_MEDIAN_MID];         // 5 样本中位 = 排序后第 2 位 / Median of five

END_METHOD

(* ---- FB_DL_CtdEx.st ---- *)
(*==============================================================================
 * 组件名称 (Component)  : FB_DL_CtdEx
 * 所属子库 (Sublibrary) : DL_Base
 * 当前版本 (Version)    : 1.0.0
 * 兼容性   (Platform)   : CODESYS 3.5 / TwinCAT 3 / 汇川 InoProShop / Machine Expert
 *                         仅依赖 Standard.library（R_TRIG），计数本体为库内显式
 *                         判界加减法（重实现最小化：仅一圈判界 + 减 1）
 * 功能描述 (Function)   : 减计数器防御包装。内部以 R_TRIG 标准实例产计数脉冲，
 *                         计数本体采用显式判界减法实现 CV 下限饱和不回绕（达
 *                         DINT 下限锁定并置诊断码）；装载优先级 bLOAD > bCD，
 *                         LOAD 按 IEC 标准语义为电平装载（CV := PV）。
 * 溯源     (Origin)     : IEC 61131-3 标准语义的道莅防御性实现
 *                         （接口语义由 IEC 61131-3 定义，clean-room 重写，
 *                         参考公开标准条款）
 * 码位     (Diag Codes) : 信息级占用区间 16#0001_0154（本件独占，仅此一码，
 *                         双事件共用一类码）
 *                         16#0001_0154 = nPV 为负值已钳 0 ／ CV 达 DINT 下限
 *                         饱和锁定（信息级，饱和是正常防御行为，不置故障）
 * 类型裁定 (Type Note)  : 码位段 16#0001_xxxx 为全库共享 32 位段，WORD 容量不足，
 *                         故 uDiag 采用 UDINT 承载（与库内 uErrorId : UDINT 惯例一致）
 * 依赖     (Depends)    : 无 DL_ 内部依赖；Standard.library: R_TRIG
 * 红线自检 (Redline)    : R1 ✓ 零全局变量与外部变量引用 ｜ R2 ✓ 零物理 IO 地址直写
 *                         R3 ✓ 纯 IEC 61131-3 ｜ R4 ✓ PV 钳位+DINT 下限判界防回绕
 *                         R5 ✓ 全变量中英双语同行注释 ｜ R6 N/A（无顺序状态机，见下）
 *                         R7 ✓ R_TRIG 实例主体无条件周期刷新
 * 说明     (Note)       : R6 标注 N/A —— 本组件为「装载/计数」双态时序逻辑，
 *                         非顺序步进状态机，无 CASE 可写；两态互斥由优先级链
 *                         （装载 > 计数）显式保证，以本节说明替代 ELSE 兜底，
 *                         符合"无状态机则标注 N/A"口径。
 * 防御行为声明 (Defense): ① nPV < 0 时钳位为 0 并置信息码 16#0001_0154
 *                           （装载后 CV=0，bQ 立即 TRUE，属组态错误提示）；
 *                         ② 下溢饱和不回绕：CV 达 DINT 下限 -2147483648 后停止
 *                           递减、保持不变并置信息码（与标准 CTD 的 DINT 回绕
 *                           行为差异点，饱和是正常防御行为）；
 *                         ③ LOAD 语义按 IEC 标准：bLOAD 为电平有效，有效期间
 *                           CV 每拍装载为钳位后 PV（非沿触发），优先级高于
 *                           bCD 计数脉冲；
 *                         ④ CV 允许为负数并继续递减至 DINT 下限（IEC CTD 标准
 *                           语义 Q = CV <= 0），下限饱和仅拦截 DINT 回绕；
 *                         ⑤ 内部状态量写入点排序审计（历史教训⑦）：PV 钳位段
 *                           与计数段对 uDiag 只写同一码值 16#0001_0154，不存在
 *                           复位类与置位类竞态，排序安全；
 *                         ⑥ DINT 下限提为只读常量 nDintMin，禁魔法数。
 * 修订历史 (Revision)   :
 *   2026-11-16  v1.0.0  首版入库（R14 批 2 · T0 快车道）
 *============================================================================*)
FUNCTION_BLOCK FB_DL_CtdEx
VAR_INPUT
    bCD   : BOOL;  // 减计数脉冲输入（内部 R_TRIG 取沿） / Count-down pulse input (edge taken by internal R_TRIG)
    bLOAD : BOOL;  // 装载输入（电平，优先级最高），CV := 钳位后 PV / Load input (level, highest priority), CV := clamped PV
    nPV   : INT;   // 预置装载值 [个]，负值将被钳位为 0 / Preset load value [count], negative values are clamped to 0
END_VAR
VAR_OUTPUT
    nCV   : DINT;   // 当前计数值 [个]，可为负，达下限饱和不回绕 / Current count [count], may go negative, saturates at lower limit without wrap
    bQ    : BOOL;   // 计数到零输出，nCV <= 0 时 TRUE / Zero-reached output, TRUE when nCV <= 0
    uDiag : UDINT;  // 诊断字，16#0001_0154=nPV 负钳 0 或 CV 下限饱和，0=无事件 / Diag word, 16#0001_0154=negative nPV clamped or CV lower saturation, 0=no event
END_VAR
VAR
    fbCdTrig  : R_TRIG;  // 内建上升沿实例，产计数脉冲 / Built-in R_TRIG instance, generates the count pulse
    nPVClamp  : DINT;    // 钳位后的预置装载值 [个]，用于装载与组态提示 / Clamped preset load value [count], used for loading and config hint
    nDintMin  : DINT := -2147483648;  // DINT 下限常量（只读语义，主体禁写）/ DINT lower-limit constant (read-only semantics, never written in body)
    xInit     : BOOL;    // 首扫初始化标志，FALSE=尚未完成上电初始化 / First-scan init flag, FALSE = power-on init not yet done
END_VAR

(*------------------------------------------------------------------------------
 * 段 1｜首扫初始化（历史教训④口径）：置于逻辑最前，首扫 CV=0、bQ=TRUE
 *      （IEC CTD 标准语义 CV<=0，首扫 0 值天然满足，非假触发）
 *      First-scan init (lesson 4): CV=0 and bQ=TRUE on first scan per IEC CTD
 *      semantics CV<=0, a natural zero value, not a false trigger
 *-----------------------------------------------------------------------------*)
IF NOT xInit THEN
    xInit    := TRUE;    // 置初始化完成标志 / Mark init as done
    nCV      := 0;       // 首扫计数值清零 [个] / Zero count on first scan [count]
    nPVClamp := 0;       // 首扫钳位预置清零 [个] / Zero clamped preset on first scan [count]
    uDiag    := 16#0000_0000;  // 首扫诊断字清零 / Clear diag word on first scan
END_IF

(*------------------------------------------------------------------------------
 * 段 2｜PV 域校验与钳位（历史教训⑨）：nPV 负值钳 0 并置信息码
 *      PV domain check and clamp (lesson 9): negative nPV clamped to 0 with code
 *-----------------------------------------------------------------------------*)
IF nPV < 0 THEN
    nPVClamp := 0;            // 负预置钳位为 0 [个] / Clamp negative preset to 0 [count]
    uDiag    := 16#0001_0154;  // 信息码：nPV 负值已钳 0 / Informational: negative nPV clamped to 0
ELSE
    nPVClamp := nPV;          // 域内直通 [个] / In-domain pass-through [count]
    uDiag    := 16#0000_0000;  // 无诊断事件，清码 / No diag event, clear code
END_IF

(*------------------------------------------------------------------------------
 * 段 3｜无条件刷新区（红线 R7）：R_TRIG 实例严禁进入任何 IF / CASE 分支
 *      Unconditional refresh zone (red line R7): no instance call inside IF / CASE
 *-----------------------------------------------------------------------------*)
fbCdTrig(CLK := bCD);  // 每扫描周期无条件取 bCD 上升沿 / Take bCD rising edge unconditionally every scan

(*------------------------------------------------------------------------------
 * 段 4｜计数主体（优先级链 bLOAD > bCD）：装载电平优先，计数沿次之；
 *      LOAD 为 IEC 标准电平装载语义（CV := PV）；下溢判界先行——CV 达 DINT
 *      下限停止递减并置饱和码，绝不回绕
 *      Count body (priority chain bLOAD > bCD): load level first, count edge
 *      second; LOAD is the IEC level-load semantics (CV := PV); underflow
 *      boundary checked before decrement, no wrap ever
 *-----------------------------------------------------------------------------*)
IF bLOAD THEN
    nCV := nPVClamp;  // 电平装载：CV := 钳位后预置值 [个] / Level load: CV := clamped preset [count]
ELSIF fbCdTrig.Q THEN
    IF nCV > nDintMin THEN
        nCV := nCV - 1;           // 域内递减 1 [个] / In-domain decrement by 1 [count]
    ELSE
        uDiag := 16#0001_0154;    // 信息码：CV 下限饱和锁定，不回绕 / Informational: CV lower-limit saturation, no wrap
    END_IF
END_IF

(*------------------------------------------------------------------------------
 * 段 5｜比较输出：按 IEC CTD 标准语义 Q = CV <= 0
 *      Compare output: per IEC CTD standard semantics Q = CV <= 0
 *-----------------------------------------------------------------------------*)
bQ := (nCV <= 0);  // 计数到零比较 [个] / Zero-reached comparison [count]
END_FUNCTION_BLOCK
